(* IEC 61131-3 sources: deprecated-refusr-repo/GP/Main/samples (part 23) *)

(* ---- RND-EXPR_roust-surfs-pairs.st ---- *)
(*
This code implements a randomly grown symbolic expression:

xor(xor(!(xor(xor(IN32, (!(!((IN49 | (!(IN19))) & (!(IN28 & (xor(xor(IN18, IN20), IN24))))))) & ((xor(xor(IN13, IN1), !(xor(xor(xor(xor(!(IN32), IN20 & IN18), IN50 & IN1), (IN10 & IN17) & (IN11 & IN39)), true & IN1)))) | (xor(xor((!(IN35)) | IN42, !(IN44 | ((!(IN28)) | IN34))), (!((xor(xor(IN28, IN8), IN8)) & IN14)) | (!(xor(xor(xor(xor(IN16, IN9), IN43), xor(xor(IN30, IN9), IN40)), IN50 | IN28))))))), xor(xor((xor(xor(!(((!(IN18)) & (!(IN40))) & (IN28 & (!(IN19)))), IN7), (!((xor(xor(IN34, IN23), IN2)) & (xor(xor(IN27, IN44), IN31)))) | (!(xor(xor(!(IN25), IN8 & IN22), IN9))))) & (xor(xor(IN3, (!(IN42)) & (xor(xor(xor(xor(IN29 & IN50, IN38 | IN40), !(IN36)), IN40), (!(IN24)) & false))), (((!(IN11)) | (!(IN14))) | ((!(IN10)) | (IN36 & IN47))) | IN15)), (!(!(IN45))) & (xor(xor(IN31 | true, IN38), xor(xor(IN43, xor(xor(IN1, (IN12 & IN45) | (IN48 | IN6)), xor(xor(xor(xor(IN28, IN15), IN16), IN6), !(IN49)))), IN13 | ((xor(xor(IN45, IN5), IN32)) & (xor(xor(IN49, IN26), IN28))))))), !((!(IN43)) | (IN45 | (IN20 & (!(xor(xor(IN16, IN7), IN9))))))))), xor(xor((IN15 & ((!(xor(xor(!(xor(xor(IN18 | IN27, xor(xor(IN38, IN31), IN37)), !(IN3))), IN8 & (!(IN28 | IN17))), (xor(xor(IN17 | IN48, xor(xor(IN42, true), true)), IN31 | IN45)) | (IN25 | (!(IN12)))))) | ((!((xor(xor(!(IN16), IN16), xor(xor(IN32, IN22), IN35))) | IN22)) & ((!(xor(xor(IN8, xor(xor(IN18, IN44), IN32)), IN10 | IN3))) & (IN48 & (IN40 | (IN42 & IN27))))))) & IN10, ((!(!(xor(xor(IN3, IN47), (!(IN36 & IN49)) | ((xor(xor(IN42, IN21), IN34)) | (xor(xor(IN24, IN27), IN13))))))) | ((!(IN3)) & IN11)) & (!(((xor(xor(IN31 & IN15, ((!(IN49)) & (xor(xor(IN42, IN39), IN29))) & IN5), (IN7 | (IN32 | IN49)) & ((!(IN32)) | IN44))) & (!(!(!(IN47 & IN34))))) | (((true | (xor(xor(!(IN5), IN9 | IN38), !(IN46)))) | (!((IN37 | IN29) | (IN12 & IN37)))) | IN9)))), !((xor(xor(xor(xor(!(IN20), IN29 | IN30), (xor(xor(IN2, (IN21 & IN3) | (IN13 | IN7)), IN28)) | (xor(xor(IN44, IN21), (!(IN49)) & (!(IN44))))), xor(xor(xor(xor(xor(xor((!(IN48)) & (xor(xor(IN4, IN4), IN39)), (IN31 & IN45) & (IN44 | IN11)), IN5), IN42 & IN13), xor(xor(IN42, (xor(xor(IN14, IN11), IN43)) & IN1), true & (!(IN29)))), !(IN20)), true | (((xor(xor(IN15, IN17), IN17)) | IN20) | (!(!(IN29)))))), (!(IN1 | (xor(xor(IN14 & IN10, !(IN14)), IN21 & IN34)))) & IN17)) | ((IN1 & (xor(xor((!(IN2 & IN15)) | IN22, (!(IN21)) | (IN15 & IN29)), !(xor(xor(IN40, IN7 & IN9), IN31))))) & (((((IN44 & IN35) & (!(IN27))) | IN14) & (IN31 | ((!(IN25)) | (!(IN45))))) | (IN34 | (!((IN22 | IN16) & IN33)))))))), !(IN31 & ((!(xor(xor(((xor(xor(IN2 & IN9, IN28 & IN31), !(IN12))) | ((IN37 | IN35) | IN39)) | ((xor(xor(IN39 & IN49, IN2), IN26 | IN19)) | IN2), xor(xor((IN41 & (!(IN16))) & (xor(xor(!(IN33), IN12 & IN24), IN29 & IN35)), ((IN50 | IN17) & (IN41 & IN40)) | IN5), xor(xor(true, xor(xor(!(IN50), xor(xor(IN37, IN38), IN12)), !(IN47))), !(IN11 | IN42)))), IN42 | IN28))) | ((IN38 & IN43) & IN36))))

*)

FUNCTION_BLOCK F_CollectInput
  VAR_IN_OUT
      Data : ARRAY[1..50] OF BOOL;
  END_VAR
  VAR_INPUT
      TICK  : BOOL := 0;
      IN1   : BOOL := 0;
      IN2   : BOOL := 0;
      IN3   : BOOL := 0;
      IN4   : BOOL := 0;
      IN5   : BOOL := 0;
      RESET : BOOL := FALSE;
  END_VAR
  VAR_OUTPUT
      Finished : BOOL;
  END_VAR
  VAR
      j    : USINT := 1;
      tock : BOOL  := 0;
  END_VAR
  IF NOT RESET AND tock = NOT TICK THEN
      Data[j]   := IN1;
      Data[j+1] := IN2;
      Data[j+2] := IN3;
      Data[j+3] := IN4;
      Data[j+4] := IN5;
      j := j + 5;
      tock := TICK;
  ELSE
      j := 1;
      tock := 0;
  END_IF;
  Finished := (j > 50);
END_FUNCTION_BLOCK

PROGRAM Boiler
  VAR
    Data  : ARRAY[1..50] OF BOOL;
    Ready : BOOL;
    CollectInput : F_CollectInput;
  END_VAR
  VAR
    TICK     AT %IX1.0 : BOOL;
    IN1      AT %IX0.3 : BOOL;
    IN2      AT %IX0.4 : BOOL;
    IN3      AT %IX0.5 : BOOL;
    IN4      AT %IX0.6 : BOOL;
    IN5      AT %IX0.7 : BOOL;
    OutReady AT %QX0.0 : BOOL := FALSE;
    FeedNext AT %QX0.1 : BOOL := FALSE;
    Out      AT %QX0.2 : BOOL;
  END_VAR
  CollectInput(TICK:=TICK, IN1:=IN1, IN2:=IN2, IN3:=IN3, IN4:=IN4, IN5:=IN5);
  Ready := CollectInput.Finished;
  FeedNext := 1;
  IF Ready THEN
    Out := (((NOT ((Data[32] XOR ((NOT (NOT ((Data[49] OR (NOT Data[19])) AND (NOT (Data[28] AND ((Data[18] XOR Data[20]) XOR Data[24])))))) AND (((Data[13] XOR Data[1]) XOR (NOT (((((NOT Data[32]) XOR (Data[20] AND Data[18])) XOR (Data[50] AND Data[1])) XOR ((Data[10] AND Data[17]) AND (Data[11] AND Data[39]))) XOR (TRUE AND Data[1])))) OR ((((NOT Data[35]) OR Data[42]) XOR (NOT (Data[44] OR ((NOT Data[28]) OR Data[34])))) XOR ((NOT (((Data[28] XOR Data[8]) XOR Data[8]) AND Data[14])) OR (NOT ((((Data[16] XOR Data[9]) XOR Data[43]) XOR ((Data[30] XOR Data[9]) XOR Data[40])) XOR (Data[50] OR Data[28])))))))) XOR ((((((NOT (((NOT Data[18]) AND (NOT Data[40])) AND (Data[28] AND (NOT Data[19])))) XOR Data[7]) XOR ((NOT (((Data[34] XOR Data[23]) XOR Data[2]) AND ((Data[27] XOR Data[44]) XOR Data[31]))) OR (NOT (((NOT Data[25]) XOR (Data[8] AND Data[22])) XOR Data[9])))) AND ((Data[3] XOR ((NOT Data[42]) AND (((((Data[29] AND Data[50]) XOR (Data[38] OR Data[40])) XOR (NOT Data[36])) XOR Data[40]) XOR ((NOT Data[24]) AND FALSE)))) XOR ((((NOT Data[11]) OR (NOT Data[14])) OR ((NOT Data[10]) OR (Data[36] AND Data[47]))) OR Data[15]))) XOR ((NOT (NOT Data[45])) AND (((Data[31] OR TRUE) XOR Data[38]) XOR ((Data[43] XOR ((Data[1] XOR ((Data[12] AND Data[45]) OR (Data[48] OR Data[6]))) XOR ((((Data[28] XOR Data[15]) XOR Data[16]) XOR Data[6]) XOR (NOT Data[49])))) XOR (Data[13] OR (((Data[45] XOR Data[5]) XOR Data[32]) AND ((Data[49] XOR Data[26]) XOR Data[28]))))))) XOR (NOT ((NOT Data[43]) OR (Data[45] OR (Data[20] AND (NOT ((Data[16] XOR Data[7]) XOR Data[9]))))))))) XOR ((((Data[15] AND ((NOT (((NOT (((Data[18] OR Data[27]) XOR ((Data[38] XOR Data[31]) XOR Data[37])) XOR (NOT Data[3]))) XOR (Data[8] AND (NOT (Data[28] OR Data[17])))) XOR ((((Data[17] OR Data[48]) XOR ((Data[42] XOR TRUE) XOR TRUE)) XOR (Data[31] OR Data[45])) OR (Data[25] OR (NOT Data[12]))))) OR ((NOT ((((NOT Data[16]) XOR Data[16]) XOR ((Data[32] XOR Data[22]) XOR Data[35])) OR Data[22])) AND ((NOT ((Data[8] XOR ((Data[18] XOR Data[44]) XOR Data[32])) XOR (Data[10] OR Data[3]))) AND (Data[48] AND (Data[40] OR (Data[42] AND Data[27]))))))) AND Data[10]) XOR (((NOT (NOT ((Data[3] XOR Data[47]) XOR ((NOT (Data[36] AND Data[49])) OR (((Data[42] XOR Data[21]) XOR Data[34]) OR ((Data[24] XOR Data[27]) XOR Data[13])))))) OR ((NOT Data[3]) AND Data[11])) AND (NOT (((((Data[31] AND Data[15]) XOR (((NOT Data[49]) AND ((Data[42] XOR Data[39]) XOR Data[29])) AND Data[5])) XOR ((Data[7] OR (Data[32] OR Data[49])) AND ((NOT Data[32]) OR Data[44]))) AND (NOT (NOT (NOT (Data[47] AND Data[34]))))) OR (((TRUE OR (((NOT Data[5]) XOR (Data[9] OR Data[38])) XOR (NOT Data[46]))) OR (NOT ((Data[37] OR Data[29]) OR (Data[12] AND Data[37])))) OR Data[9]))))) XOR (NOT ((((((NOT Data[20]) XOR (Data[29] OR Data[30])) XOR (((Data[2] XOR ((Data[21] AND Data[3]) OR (Data[13] OR Data[7]))) XOR Data[28]) OR ((Data[44] XOR Data[21]) XOR ((NOT Data[49]) AND (NOT Data[44]))))) XOR ((((((((NOT Data[48]) AND ((Data[4] XOR Data[4]) XOR Data[39])) XOR ((Data[31] AND Data[45]) AND (Data[44] OR Data[11]))) XOR Data[5]) XOR (Data[42] AND Data[13])) XOR ((Data[42] XOR (((Data[14] XOR Data[11]) XOR Data[43]) AND Data[1])) XOR (TRUE AND (NOT Data[29])))) XOR (NOT Data[20])) XOR (TRUE OR ((((Data[15] XOR Data[17]) XOR Data[17]) OR Data[20]) OR (NOT (NOT Data[29])))))) XOR ((NOT (Data[1] OR (((Data[14] AND Data[10]) XOR (NOT Data[14])) XOR (Data[21] AND Data[34])))) AND Data[17])) OR ((Data[1] AND ((((NOT (Data[2] AND Data[15])) OR Data[22]) XOR ((NOT Data[21]) OR (Data[15] AND Data[29]))) XOR (NOT ((Data[40] XOR (Data[7] AND Data[9])) XOR Data[31])))) AND (((((Data[44] AND Data[35]) AND (NOT Data[27])) OR Data[14]) AND (Data[31] OR ((NOT Data[25]) OR (NOT Data[45])))) OR (Data[34] OR (NOT ((Data[22] OR Data[16]) AND Data[33]))))))))) XOR (NOT (Data[31] AND ((NOT (((((((Data[2] AND Data[9]) XOR (Data[28] AND Data[31])) XOR (NOT Data[12])) OR ((Data[37] OR Data[35]) OR Data[39])) OR ((((Data[39] AND Data[49]) XOR Data[2]) XOR (Data[26] OR Data[19])) OR Data[2])) XOR ((((Data[41] AND (NOT Data[16])) AND (((NOT Data[33]) XOR (Data[12] AND Data[24])) XOR (Data[29] AND Data[35]))) XOR (((Data[50] OR Data[17]) AND (Data[41] AND Data[40])) OR Data[5])) XOR ((TRUE XOR (((NOT Data[50]) XOR ((Data[37] XOR Data[38]) XOR Data[12])) XOR (NOT Data[47]))) XOR (NOT (Data[11] OR Data[42]))))) XOR (Data[42] OR Data[28]))) OR ((Data[38] AND Data[43]) AND Data[36])))));
    OutReady := 1;
    CollectInput(RESET:=TRUE);
  END_IF;
END_PROGRAM

CONFIGURATION Config0
  RESOURCE Res0 ON PLC
    TASK task0(INTERVAL := T#20ms,PRIORITY := 0);
    PROGRAM instance0 WITH task0 : Boiler;
  END_RESOURCE
END_CONFIGURATION

(* ---- RND-EXPR_sepal-sighs-minis.st ---- *)
(*
This code implements a randomly grown symbolic expression:

((xor(xor(!(IN17), IN3), IN42 & (!(!((!(xor(xor(IN42 & IN8, IN18), IN49))) | (!(IN32))))))) & ((!(!((IN47 | (IN12 & (xor(xor(!(IN9), IN41 & IN17), IN45)))) & (xor(xor(IN6 & (IN23 | (IN31 | IN44)), xor(xor((!(IN32)) & (!(IN23)), IN42 & (IN50 | IN34)), xor(xor(!(IN34), !(IN32)), IN15))), xor(xor(IN33, xor(xor(IN45 & IN5, IN11 & IN16), IN3 | IN4)), !(!(IN15)))))))) & (((xor(xor(((xor(xor(IN50 | IN14, IN46 & IN40), xor(xor(IN3, IN41), IN9))) & (IN22 & IN28)) | (xor(xor(IN41 | (IN26 & IN10), xor(xor(IN42 & IN12, xor(xor(IN32, IN46), IN35)), IN1 & IN11)), xor(xor(xor(xor(IN43, IN19), IN38), IN27 | IN21), !(IN10)))), !(xor(xor((xor(xor(IN7, IN50), IN1)) | IN6, (IN35 & IN3) | (!(IN28))), xor(xor(IN7 & IN16, IN37 | IN33), IN11)))), (!((!(IN25)) | (!(IN41)))) & ((!(IN33 & true)) & (!(!(IN5)))))) & (xor(xor(IN12, !(IN17)), (((!(IN28)) & (xor(xor(IN4, IN22), IN12))) | ((IN4 & IN38) & IN37)) | true))) | IN6))) & (xor(xor(!(IN24), xor(xor(!((xor(xor(IN48 | (!((IN17 & IN14) | IN31)), (xor(xor(true, xor(xor(xor(xor(IN16, IN16), IN17), !(IN23)), IN2)), (!(IN45)) | (xor(xor(IN31, IN48), IN25)))) & (!(xor(xor(IN6, IN41 & IN37), IN38)))), (IN26 | ((IN7 & IN2) | (IN17 | false))) & (xor(xor(IN42 & (IN28 | IN44), (IN16 & IN26) | (IN21 | IN13)), (IN11 & IN4) | (IN48 | IN47))))) & ((!(false & ((xor(xor(IN20, IN8), IN2)) | (IN36 & IN18)))) & IN47)), xor(xor(((false & (xor(xor(xor(xor(IN27 | IN30, xor(xor(IN23, IN27), IN7)), IN21), !(IN50)), (!(IN35)) & (xor(xor(IN21, IN7), IN17))))) | ((((IN9 | IN5) | (xor(xor(IN46, IN31), IN33))) | IN14) | IN32)) | (((!(IN19)) & IN21) & (!((!(IN44 & IN26)) | IN42))), xor(xor(!(IN34), (IN31 | (xor(xor(IN20, IN9), IN30))) | (xor(xor(IN21, xor(xor((IN29 | IN5) | (IN10 & IN14), xor(xor(IN41 & IN34, xor(xor(IN20, IN4), IN29)), IN29 & IN17)), IN39 | (IN7 & IN43))), ((!(IN40)) | IN50) | (!(IN17))))), xor(xor(xor(xor(IN31, IN24), ((IN30 | IN5) & (!(IN48))) | ((xor(xor(IN16, IN13), IN34)) & (!(IN16)))), (xor(xor(IN29 | IN25, xor(xor(xor(xor(IN20, IN40), IN9), IN26 | IN20), IN43 | IN32)), (xor(xor(IN35, IN6), IN33)) | (IN30 | IN7))) & (((true | IN15) | (IN46 | IN5)) | ((xor(xor(IN20, IN39), IN5)) | (IN48 | IN20)))), ((!(IN11 & IN1)) | ((xor(xor(IN5, IN25), IN49)) | (IN3 & IN43))) | (!(xor(xor(IN22, xor(xor(IN40, IN26), IN7)), xor(xor(IN10, IN10), IN44))))))), !(xor(xor(!(xor(xor((!(IN32)) | (xor(xor(IN28, IN4), IN11)), (IN7 | IN49) & (IN19 | IN17)), xor(xor(xor(xor(IN50, IN4), IN7), !(IN25)), !(IN10)))), (xor(xor(IN18 & (IN23 | IN36), xor(xor(IN36 | false, IN31 | IN19), IN15 & IN5)), !(IN41))) | (!(!(xor(xor(IN34, IN8), true))))), IN10 & (((IN39 & IN8) | (xor(xor(IN37, IN1), IN46))) | ((xor(xor(IN21, IN1), IN16)) | (false | IN1))))))), IN25 & (IN31 & (IN20 & IN46)))), IN38 | (!(IN32))))

*)

FUNCTION_BLOCK F_CollectInput
  VAR_IN_OUT
      Data : ARRAY[1..50] OF BOOL;
  END_VAR
  VAR_INPUT
      TICK  : BOOL := 0;
      IN1   : BOOL := 0;
      IN2   : BOOL := 0;
      IN3   : BOOL := 0;
      IN4   : BOOL := 0;
      IN5   : BOOL := 0;
      RESET : BOOL := FALSE;
  END_VAR
  VAR_OUTPUT
      Finished : BOOL;
  END_VAR
  VAR
      j    : USINT := 1;
      tock : BOOL  := 0;
  END_VAR
  IF NOT RESET AND tock = NOT TICK THEN
      Data[j]   := IN1;
      Data[j+1] := IN2;
      Data[j+2] := IN3;
      Data[j+3] := IN4;
      Data[j+4] := IN5;
      j := j + 5;
      tock := TICK;
  ELSE
      j := 1;
      tock := 0;
  END_IF;
  Finished := (j > 50);
END_FUNCTION_BLOCK

PROGRAM Boiler
  VAR
    Data  : ARRAY[1..50] OF BOOL;
    Ready : BOOL;
    CollectInput : F_CollectInput;
  END_VAR
  VAR
    TICK     AT %IX1.0 : BOOL;
    IN1      AT %IX0.3 : BOOL;
    IN2      AT %IX0.4 : BOOL;
    IN3      AT %IX0.5 : BOOL;
    IN4      AT %IX0.6 : BOOL;
    IN5      AT %IX0.7 : BOOL;
    OutReady AT %QX0.0 : BOOL := FALSE;
    FeedNext AT %QX0.1 : BOOL := FALSE;
    Out      AT %QX0.2 : BOOL;
  END_VAR
  CollectInput(TICK:=TICK, IN1:=IN1, IN2:=IN2, IN3:=IN3, IN4:=IN4, IN5:=IN5);
  Ready := CollectInput.Finished;
  FeedNext := 1;
  IF Ready THEN
    Out := (((((NOT Data[17]) XOR Data[3]) XOR (Data[42] AND (NOT (NOT ((NOT (((Data[42] AND Data[8]) XOR Data[18]) XOR Data[49])) OR (NOT Data[32])))))) AND ((NOT (NOT ((Data[47] OR (Data[12] AND (((NOT Data[9]) XOR (Data[41] AND Data[17])) XOR Data[45]))) AND (((Data[6] AND (Data[23] OR (Data[31] OR Data[44]))) XOR ((((NOT Data[32]) AND (NOT Data[23])) XOR (Data[42] AND (Data[50] OR Data[34]))) XOR (((NOT Data[34]) XOR (NOT Data[32])) XOR Data[15]))) XOR ((Data[33] XOR (((Data[45] AND Data[5]) XOR (Data[11] AND Data[16])) XOR (Data[3] OR Data[4]))) XOR (NOT (NOT Data[15]))))))) AND (((((((((Data[50] OR Data[14]) XOR (Data[46] AND Data[40])) XOR ((Data[3] XOR Data[41]) XOR Data[9])) AND (Data[22] AND Data[28])) OR (((Data[41] OR (Data[26] AND Data[10])) XOR (((Data[42] AND Data[12]) XOR ((Data[32] XOR Data[46]) XOR Data[35])) XOR (Data[1] AND Data[11]))) XOR ((((Data[43] XOR Data[19]) XOR Data[38]) XOR (Data[27] OR Data[21])) XOR (NOT Data[10])))) XOR (NOT (((((Data[7] XOR Data[50]) XOR Data[1]) OR Data[6]) XOR ((Data[35] AND Data[3]) OR (NOT Data[28]))) XOR (((Data[7] AND Data[16]) XOR (Data[37] OR Data[33])) XOR Data[11])))) XOR ((NOT ((NOT Data[25]) OR (NOT Data[41]))) AND ((NOT (Data[33] AND TRUE)) AND (NOT (NOT Data[5]))))) AND ((Data[12] XOR (NOT Data[17])) XOR ((((NOT Data[28]) AND ((Data[4] XOR Data[22]) XOR Data[12])) OR ((Data[4] AND Data[38]) AND Data[37])) OR TRUE))) OR Data[6]))) AND (((NOT Data[24]) XOR (((NOT ((((Data[48] OR (NOT ((Data[17] AND Data[14]) OR Data[31]))) XOR (((TRUE XOR ((((Data[16] XOR Data[16]) XOR Data[17]) XOR (NOT Data[23])) XOR Data[2])) XOR ((NOT Data[45]) OR ((Data[31] XOR Data[48]) XOR Data[25]))) AND (NOT ((Data[6] XOR (Data[41] AND Data[37])) XOR Data[38])))) XOR ((Data[26] OR ((Data[7] AND Data[2]) OR (Data[17] OR FALSE))) AND (((Data[42] AND (Data[28] OR Data[44])) XOR ((Data[16] AND Data[26]) OR (Data[21] OR Data[13]))) XOR ((Data[11] AND Data[4]) OR (Data[48] OR Data[47]))))) AND ((NOT (FALSE AND (((Data[20] XOR Data[8]) XOR Data[2]) OR (Data[36] AND Data[18])))) AND Data[47]))) XOR (((((FALSE AND (((((Data[27] OR Data[30]) XOR ((Data[23] XOR Data[27]) XOR Data[7])) XOR Data[21]) XOR (NOT Data[50])) XOR ((NOT Data[35]) AND ((Data[21] XOR Data[7]) XOR Data[17])))) OR ((((Data[9] OR Data[5]) OR ((Data[46] XOR Data[31]) XOR Data[33])) OR Data[14]) OR Data[32])) OR (((NOT Data[19]) AND Data[21]) AND (NOT ((NOT (Data[44] AND Data[26])) OR Data[42])))) XOR (((NOT Data[34]) XOR ((Data[31] OR ((Data[20] XOR Data[9]) XOR Data[30])) OR ((Data[21] XOR ((((Data[29] OR Data[5]) OR (Data[10] AND Data[14])) XOR (((Data[41] AND Data[34]) XOR ((Data[20] XOR Data[4]) XOR Data[29])) XOR (Data[29] AND Data[17]))) XOR (Data[39] OR (Data[7] AND Data[43])))) XOR (((NOT Data[40]) OR Data[50]) OR (NOT Data[17]))))) XOR ((((Data[31] XOR Data[24]) XOR (((Data[30] OR Data[5]) AND (NOT Data[48])) OR (((Data[16] XOR Data[13]) XOR Data[34]) AND (NOT Data[16])))) XOR ((((Data[29] OR Data[25]) XOR ((((Data[20] XOR Data[40]) XOR Data[9]) XOR (Data[26] OR Data[20])) XOR (Data[43] OR Data[32]))) XOR (((Data[35] XOR Data[6]) XOR Data[33]) OR (Data[30] OR Data[7]))) AND (((TRUE OR Data[15]) OR (Data[46] OR Data[5])) OR (((Data[20] XOR Data[39]) XOR Data[5]) OR (Data[48] OR Data[20]))))) XOR (((NOT (Data[11] AND Data[1])) OR (((Data[5] XOR Data[25]) XOR Data[49]) OR (Data[3] AND Data[43]))) OR (NOT ((Data[22] XOR ((Data[40] XOR Data[26]) XOR Data[7])) XOR ((Data[10] XOR Data[10]) XOR Data[44]))))))) XOR (NOT (((NOT ((((NOT Data[32]) OR ((Data[28] XOR Data[4]) XOR Data[11])) XOR ((Data[7] OR Data[49]) AND (Data[19] OR Data[17]))) XOR ((((Data[50] XOR Data[4]) XOR Data[7]) XOR (NOT Data[25])) XOR (NOT Data[10])))) XOR ((((Data[18] AND (Data[23] OR Data[36])) XOR (((Data[36] OR FALSE) XOR (Data[31] OR Data[19])) XOR (Data[15] AND Data[5]))) XOR (NOT Data[41])) OR (NOT (NOT ((Data[34] XOR Data[8]) XOR TRUE))))) XOR (Data[10] AND (((Data[39] AND Data[8]) OR ((Data[37] XOR Data[1]) XOR Data[46])) OR (((Data[21] XOR Data[1]) XOR Data[16]) OR (FALSE OR Data[1])))))))) XOR (Data[25] AND (Data[31] AND (Data[20] AND Data[46]))))) XOR (Data[38] OR (NOT Data[32]))));
    OutReady := 1;
    CollectInput(RESET:=TRUE);
  END_IF;
END_PROGRAM

CONFIGURATION Config0
  RESOURCE Res0 ON PLC
    TASK task0(INTERVAL := T#20ms,PRIORITY := 0);
    PROGRAM instance0 WITH task0 : Boiler;
  END_RESOURCE
END_CONFIGURATION

(* ---- RND-EXPR_sewed-hokey-cooch.st ---- *)
(*
This code implements a randomly grown symbolic expression:

!(((!(IN1)) | (xor(xor(!(IN4 | (!(xor(xor((!(IN21)) | (IN10 | IN34), (IN32 & IN39) & (xor(xor(IN33, IN21), IN30))), !(IN10 & IN16))))), !(!(!(xor(xor(IN12 & (!(IN27)), xor(xor(IN33 | IN30, IN41 & IN39), !(IN28))), IN32))))), xor(xor(!(!(IN49)), xor(xor((((IN3 & IN10) | (IN5 & IN27)) | IN6) & (IN43 | (xor(xor(IN8 | IN6, IN18 | IN20), IN22))), ((xor(xor(!(IN49), xor(xor(IN25, IN15), IN10)), xor(xor(IN36, IN47), IN50))) & false) | (!(xor(xor(!(IN13), IN25), xor(xor(IN8, IN43), IN45))))), IN44)), !(xor(xor(xor(xor((IN50 | IN36) | IN39, IN13), IN21), IN46 & IN31), IN9)))))) & (xor(xor(!((!(IN49)) | (xor(xor(!(IN31), IN49), (xor(xor(IN13, (xor(xor(IN6, IN49), IN32)) & (xor(xor(IN30, IN18), IN32))), IN42 | (IN13 | IN3))) & IN32))), ((!(xor(xor(xor(xor(IN31, IN16 | (!(IN20))), (true | IN11) | (IN30 & IN6)), ((xor(xor(IN5, IN18), IN47)) | (xor(xor(IN35, IN32), IN7))) & (!(IN35 | IN25))), (xor(xor(IN45 | IN27, !(IN16)), IN28 & IN24)) & ((IN12 | IN15) | (!(IN26)))))) & (!(IN14 & (((IN50 | IN36) & (!(IN18))) | (xor(xor(false, IN20 | IN26), IN25 | IN46)))))) & (!(IN16))), !((xor(xor((xor(xor((xor(xor(IN18, IN5), IN4)) & (IN10 | IN28), (IN14 | IN50) & (xor(xor(IN31, IN38), IN9))), (IN6 | IN10) | (IN46 | IN30))) | IN8, xor(xor((IN26 & (xor(xor(IN38, IN2), IN26))) & IN24, xor(xor(IN39, (xor(xor(IN4, IN26), IN46)) & (IN21 | IN23)), (IN46 | IN28) & (IN43 & IN9))), IN47)), (!((xor(xor(IN32, IN28), IN18)) & (IN11 & IN35))) & (((xor(xor(IN50, false), IN45)) & IN3) | (xor(xor(IN8, IN14 & IN13), IN48))))) | (((!(IN19)) | (IN26 & (!(!(IN22))))) & IN12)))))

*)

FUNCTION_BLOCK F_CollectInput
  VAR_IN_OUT
      Data : ARRAY[1..50] OF BOOL;
  END_VAR
  VAR_INPUT
      TICK  : BOOL := 0;
      IN1   : BOOL := 0;
      IN2   : BOOL := 0;
      IN3   : BOOL := 0;
      IN4   : BOOL := 0;
      IN5   : BOOL := 0;
      RESET : BOOL := FALSE;
  END_VAR
  VAR_OUTPUT
      Finished : BOOL;
  END_VAR
  VAR
      j    : USINT := 1;
      tock : BOOL  := 0;
  END_VAR
  IF NOT RESET AND tock = NOT TICK THEN
      Data[j]   := IN1;
      Data[j+1] := IN2;
      Data[j+2] := IN3;
      Data[j+3] := IN4;
      Data[j+4] := IN5;
      j := j + 5;
      tock := TICK;
  ELSE
      j := 1;
      tock := 0;
  END_IF;
  Finished := (j > 50);
END_FUNCTION_BLOCK

PROGRAM Boiler
  VAR
    Data  : ARRAY[1..50] OF BOOL;
    Ready : BOOL;
    CollectInput : F_CollectInput;
  END_VAR
  VAR
    TICK     AT %IX1.0 : BOOL;
    IN1      AT %IX0.3 : BOOL;
    IN2      AT %IX0.4 : BOOL;
    IN3      AT %IX0.5 : BOOL;
    IN4      AT %IX0.6 : BOOL;
    IN5      AT %IX0.7 : BOOL;
    OutReady AT %QX0.0 : BOOL := FALSE;
    FeedNext AT %QX0.1 : BOOL := FALSE;
    Out      AT %QX0.2 : BOOL;
  END_VAR
  CollectInput(TICK:=TICK, IN1:=IN1, IN2:=IN2, IN3:=IN3, IN4:=IN4, IN5:=IN5);
  Ready := CollectInput.Finished;
  FeedNext := 1;
  IF Ready THEN
    Out := (NOT (((NOT Data[1]) OR (((NOT (Data[4] OR (NOT ((((NOT Data[21]) OR (Data[10] OR Data[34])) XOR ((Data[32] AND Data[39]) AND ((Data[33] XOR Data[21]) XOR Data[30]))) XOR (NOT (Data[10] AND Data[16])))))) XOR (NOT (NOT (NOT (((Data[12] AND (NOT Data[27])) XOR (((Data[33] OR Data[30]) XOR (Data[41] AND Data[39])) XOR (NOT Data[28]))) XOR Data[32]))))) XOR (((NOT (NOT Data[49])) XOR ((((((Data[3] AND Data[10]) OR (Data[5] AND Data[27])) OR Data[6]) AND (Data[43] OR (((Data[8] OR Data[6]) XOR (Data[18] OR Data[20])) XOR Data[22]))) XOR (((((NOT Data[49]) XOR ((Data[25] XOR Data[15]) XOR Data[10])) XOR ((Data[36] XOR Data[47]) XOR Data[50])) AND FALSE) OR (NOT (((NOT Data[13]) XOR Data[25]) XOR ((Data[8] XOR Data[43]) XOR Data[45]))))) XOR Data[44])) XOR (NOT ((((((Data[50] OR Data[36]) OR Data[39]) XOR Data[13]) XOR Data[21]) XOR (Data[46] AND Data[31])) XOR Data[9]))))) AND (((NOT ((NOT Data[49]) OR (((NOT Data[31]) XOR Data[49]) XOR (((Data[13] XOR (((Data[6] XOR Data[49]) XOR Data[32]) AND ((Data[30] XOR Data[18]) XOR Data[32]))) XOR (Data[42] OR (Data[13] OR Data[3]))) AND Data[32])))) XOR (((NOT ((((Data[31] XOR (Data[16] OR (NOT Data[20]))) XOR ((TRUE OR Data[11]) OR (Data[30] AND Data[6]))) XOR ((((Data[5] XOR Data[18]) XOR Data[47]) OR ((Data[35] XOR Data[32]) XOR Data[7])) AND (NOT (Data[35] OR Data[25])))) XOR ((((Data[45] OR Data[27]) XOR (NOT Data[16])) XOR (Data[28] AND Data[24])) AND ((Data[12] OR Data[15]) OR (NOT Data[26]))))) AND (NOT (Data[14] AND (((Data[50] OR Data[36]) AND (NOT Data[18])) OR ((FALSE XOR (Data[20] OR Data[26])) XOR (Data[25] OR Data[46])))))) AND (NOT Data[16]))) XOR (NOT (((((((((Data[18] XOR Data[5]) XOR Data[4]) AND (Data[10] OR Data[28])) XOR ((Data[14] OR Data[50]) AND ((Data[31] XOR Data[38]) XOR Data[9]))) XOR ((Data[6] OR Data[10]) OR (Data[46] OR Data[30]))) OR Data[8]) XOR ((((Data[26] AND ((Data[38] XOR Data[2]) XOR Data[26])) AND Data[24]) XOR ((Data[39] XOR (((Data[4] XOR Data[26]) XOR Data[46]) AND (Data[21] OR Data[23]))) XOR ((Data[46] OR Data[28]) AND (Data[43] AND Data[9])))) XOR Data[47])) XOR ((NOT (((Data[32] XOR Data[28]) XOR Data[18]) AND (Data[11] AND Data[35]))) AND ((((Data[50] XOR FALSE) XOR Data[45]) AND Data[3]) OR ((Data[8] XOR (Data[14] AND Data[13])) XOR Data[48])))) OR (((NOT Data[19]) OR (Data[26] AND (NOT (NOT Data[22])))) AND Data[12]))))));
    OutReady := 1;
    CollectInput(RESET:=TRUE);
  END_IF;
END_PROGRAM

CONFIGURATION Config0
  RESOURCE Res0 ON PLC
    TASK task0(INTERVAL := T#20ms,PRIORITY := 0);
    PROGRAM instance0 WITH task0 : Boiler;
  END_RESOURCE
END_CONFIGURATION

(* ---- RND-EXPR_sisal-keens-dweeb.st ---- *)
(*
This code implements a randomly grown symbolic expression:

((IN8 & (xor(xor(xor(xor(((!(xor(xor(IN20 & IN27, IN16 & IN35), !(IN38)))) | (xor(xor(IN48, (xor(xor(IN13, IN11), IN50)) | (xor(xor(IN27, IN2), IN19))), xor(xor(IN10, xor(xor(IN3, IN44), IN33)), !(IN13))))) & ((((!(IN49)) | IN45) | ((xor(xor(IN37, IN11), IN42)) & (!(IN15)))) | ((IN38 & (false | IN44)) | ((xor(xor(IN48, IN7), IN31)) & (!(IN5))))), IN48), !((!(IN46)) | ((!(!(IN4))) | (!(IN23 | IN49))))), (!(xor(xor((IN49 & (!(IN6))) & IN43, xor(xor(IN45, !(IN11 & IN3)), (xor(xor(IN10, IN26), IN11)) & (IN38 & IN47))), IN10))) & ((xor(xor(xor(xor(xor(xor(IN44 | IN8, IN37), xor(xor(true, IN3), IN6)), !(IN43 & IN23)), IN6), (!(IN23 & IN33)) & (!(IN39 | IN20))), xor(xor((!(IN21)) & (IN28 | IN37), !(IN33 | IN4)), IN40))) | (!(((!(IN41)) & IN50) & ((xor(xor(IN17, IN41), IN2)) & (IN10 & IN29)))))), xor(xor(IN13, (xor(xor(!(xor(xor(!(IN25), IN30 & IN3), !(IN26))), xor(xor((IN34 | IN33) | (!(IN36)), !(IN43 | IN2)), xor(xor(IN10 & IN46, !(IN22)), xor(xor(IN44, IN37), IN16)))), xor(xor((xor(xor(IN36, IN11), IN27)) | (IN13 | IN50), (IN42 & IN34) & (IN5 & IN43)), xor(xor(IN35, !(IN35)), xor(xor(IN1, IN26), IN25))))) | (xor(xor(!(IN39), xor(xor(!(IN45 | IN21), (IN44 & IN4) & (IN15 & IN10)), !(xor(xor(IN22, IN31), IN43)))), xor(xor((xor(xor(IN15, IN44), IN15)) & (IN25 | IN26), xor(xor(IN20 & IN21, IN14 & IN13), !(IN20))), (IN50 | IN32) | (IN7 & IN7))))), (xor(xor(!((IN16 & IN46) & (xor(xor(IN50, IN17), IN23))), IN22 & ((!(IN22)) | true)), (!(xor(xor(IN30, IN23), IN12))) | (xor(xor(IN27 | IN25, xor(xor(IN32, IN20), IN47)), xor(xor(IN49, IN34), false))))) | (xor(xor(IN28, ((xor(xor(IN22, IN8), IN38)) | IN20) | (!(IN17 & IN39))), ((xor(xor(IN8, IN50), IN25)) & (IN25 & IN41)) | IN40)))))) | IN43) | (!(!(xor(xor(xor(xor(!(!(!((!(IN47)) | (xor(xor(IN48, IN32), IN40))))), xor(xor(xor(xor(IN26 & (IN36 & (IN50 | IN12)), ((IN19 & IN10) & IN42) | (xor(xor(xor(xor(IN48, IN40), IN26), IN37 & false), IN26 | IN44))), (IN23 | (IN47 | IN39)) & (xor(xor(IN31 | IN24, IN26 & IN6), !(IN11)))), !(IN22)), !(IN4))), IN18 | IN18), xor(xor(IN50, (xor(xor(xor(xor(xor(xor(IN38, IN39 | IN10), xor(xor(IN36, IN16), IN5)), !(IN43)), (xor(xor(IN43, IN20), IN44)) & (!(IN24))), ((xor(xor(IN27, IN1), IN9)) | (xor(xor(IN4, IN24), IN13))) & IN12), ((IN29 | IN47) | (!(IN32))) | IN1)) | (xor(xor(((IN41 | IN14) & (IN15 & IN9)) & IN9, (!(IN23)) | (xor(xor(IN13 | IN38, IN13), xor(xor(IN36, IN48), IN31)))), xor(xor((IN7 | IN11) | (!(IN34)), (!(IN34)) | (IN43 & IN1)), (IN49 | IN16) | (!(IN49)))))), xor(xor((((false | IN17) | (xor(xor(IN3, IN13), IN3))) | (!(IN16 & true))) | (IN1 | IN25), ((!(IN50)) & (!(IN36 & IN1))) | (!(!(xor(xor(IN48, IN46), IN35))))), xor(xor(IN19 & ((IN28 & IN49) & (IN43 | IN40)), IN14), (!(IN38 | IN6)) & IN50)))), IN48 & (xor(xor(((!(IN41)) | ((xor(xor(IN14, IN38), IN48)) & IN50)) & ((xor(xor(IN11, IN18 & IN7), IN7 | IN20)) | (IN8 & (xor(xor(IN8, IN23), IN20)))), xor(xor((xor(xor(IN26 & IN21, IN4 | IN14), xor(xor(IN31, false), IN18))) & (xor(xor(IN37, IN14 & IN47), xor(xor(IN14, IN8), IN37))), !((xor(xor(IN3, IN24), IN28)) & IN29)), (IN27 | (!(IN44))) & IN22)), (!(IN29)) | (!((!(IN36)) | (IN23 | IN34)))))))))

*)

FUNCTION_BLOCK F_CollectInput
  VAR_IN_OUT
      Data : ARRAY[1..50] OF BOOL;
  END_VAR
  VAR_INPUT
      TICK  : BOOL := 0;
      IN1   : BOOL := 0;
      IN2   : BOOL := 0;
      IN3   : BOOL := 0;
      IN4   : BOOL := 0;
      IN5   : BOOL := 0;
      RESET : BOOL := FALSE;
  END_VAR
  VAR_OUTPUT
      Finished : BOOL;
  END_VAR
  VAR
      j    : USINT := 1;
      tock : BOOL  := 0;
  END_VAR
  IF NOT RESET AND tock = NOT TICK THEN
      Data[j]   := IN1;
      Data[j+1] := IN2;
      Data[j+2] := IN3;
      Data[j+3] := IN4;
      Data[j+4] := IN5;
      j := j + 5;
      tock := TICK;
  ELSE
      j := 1;
      tock := 0;
  END_IF;
  Finished := (j > 50);
END_FUNCTION_BLOCK

PROGRAM Boiler
  VAR
    Data  : ARRAY[1..50] OF BOOL;
    Ready : BOOL;
    CollectInput : F_CollectInput;
  END_VAR
  VAR
    TICK     AT %IX1.0 : BOOL;
    IN1      AT %IX0.3 : BOOL;
    IN2      AT %IX0.4 : BOOL;
    IN3      AT %IX0.5 : BOOL;
    IN4      AT %IX0.6 : BOOL;
    IN5      AT %IX0.7 : BOOL;
    OutReady AT %QX0.0 : BOOL := FALSE;
    FeedNext AT %QX0.1 : BOOL := FALSE;
    Out      AT %QX0.2 : BOOL;
  END_VAR
  CollectInput(TICK:=TICK, IN1:=IN1, IN2:=IN2, IN3:=IN3, IN4:=IN4, IN5:=IN5);
  Ready := CollectInput.Finished;
  FeedNext := 1;
  IF Ready THEN
    Out := (((Data[8] AND (((((((NOT (((Data[20] AND Data[27]) XOR (Data[16] AND Data[35])) XOR (NOT Data[38]))) OR ((Data[48] XOR (((Data[13] XOR Data[11]) XOR Data[50]) OR ((Data[27] XOR Data[2]) XOR Data[19]))) XOR ((Data[10] XOR ((Data[3] XOR Data[44]) XOR Data[33])) XOR (NOT Data[13])))) AND ((((NOT Data[49]) OR Data[45]) OR (((Data[37] XOR Data[11]) XOR Data[42]) AND (NOT Data[15]))) OR ((Data[38] AND (FALSE OR Data[44])) OR (((Data[48] XOR Data[7]) XOR Data[31]) AND (NOT Data[5]))))) XOR Data[48]) XOR (NOT ((NOT Data[46]) OR ((NOT (NOT Data[4])) OR (NOT (Data[23] OR Data[49])))))) XOR ((NOT ((((Data[49] AND (NOT Data[6])) AND Data[43]) XOR ((Data[45] XOR (NOT (Data[11] AND Data[3]))) XOR (((Data[10] XOR Data[26]) XOR Data[11]) AND (Data[38] AND Data[47])))) XOR Data[10])) AND ((((((((Data[44] OR Data[8]) XOR Data[37]) XOR ((TRUE XOR Data[3]) XOR Data[6])) XOR (NOT (Data[43] AND Data[23]))) XOR Data[6]) XOR ((NOT (Data[23] AND Data[33])) AND (NOT (Data[39] OR Data[20])))) XOR ((((NOT Data[21]) AND (Data[28] OR Data[37])) XOR (NOT (Data[33] OR Data[4]))) XOR Data[40])) OR (NOT (((NOT Data[41]) AND Data[50]) AND (((Data[17] XOR Data[41]) XOR Data[2]) AND (Data[10] AND Data[29]))))))) XOR ((Data[13] XOR ((((NOT (((NOT Data[25]) XOR (Data[30] AND Data[3])) XOR (NOT Data[26]))) XOR ((((Data[34] OR Data[33]) OR (NOT Data[36])) XOR (NOT (Data[43] OR Data[2]))) XOR (((Data[10] AND Data[46]) XOR (NOT Data[22])) XOR ((Data[44] XOR Data[37]) XOR Data[16])))) XOR (((((Data[36] XOR Data[11]) XOR Data[27]) OR (Data[13] OR Data[50])) XOR ((Data[42] AND Data[34]) AND (Data[5] AND Data[43]))) XOR ((Data[35] XOR (NOT Data[35])) XOR ((Data[1] XOR Data[26]) XOR Data[25])))) OR (((NOT Data[39]) XOR (((NOT (Data[45] OR Data[21])) XOR ((Data[44] AND Data[4]) AND (Data[15] AND Data[10]))) XOR (NOT ((Data[22] XOR Data[31]) XOR Data[43])))) XOR (((((Data[15] XOR Data[44]) XOR Data[15]) AND (Data[25] OR Data[26])) XOR (((Data[20] AND Data[21]) XOR (Data[14] AND Data[13])) XOR (NOT Data[20]))) XOR ((Data[50] OR Data[32]) OR (Data[7] AND Data[7])))))) XOR ((((NOT ((Data[16] AND Data[46]) AND ((Data[50] XOR Data[17]) XOR Data[23]))) XOR (Data[22] AND ((NOT Data[22]) OR TRUE))) XOR ((NOT ((Data[30] XOR Data[23]) XOR Data[12])) OR (((Data[27] OR Data[25]) XOR ((Data[32] XOR Data[20]) XOR Data[47])) XOR ((Data[49] XOR Data[34]) XOR FALSE)))) OR ((Data[28] XOR ((((Data[22] XOR Data[8]) XOR Data[38]) OR Data[20]) OR (NOT (Data[17] AND Data[39])))) XOR ((((Data[8] XOR Data[50]) XOR Data[25]) AND (Data[25] AND Data[41])) OR Data[40])))))) OR Data[43]) OR (NOT (NOT (((((NOT (NOT (NOT ((NOT Data[47]) OR ((Data[48] XOR Data[32]) XOR Data[40]))))) XOR (((((Data[26] AND (Data[36] AND (Data[50] OR Data[12]))) XOR (((Data[19] AND Data[10]) AND Data[42]) OR ((((Data[48] XOR Data[40]) XOR Data[26]) XOR (Data[37] AND FALSE)) XOR (Data[26] OR Data[44])))) XOR ((Data[23] OR (Data[47] OR Data[39])) AND (((Data[31] OR Data[24]) XOR (Data[26] AND Data[6])) XOR (NOT Data[11])))) XOR (NOT Data[22])) XOR (NOT Data[4]))) XOR (Data[18] OR Data[18])) XOR ((Data[50] XOR (((((((Data[38] XOR (Data[39] OR Data[10])) XOR ((Data[36] XOR Data[16]) XOR Data[5])) XOR (NOT Data[43])) XOR (((Data[43] XOR Data[20]) XOR Data[44]) AND (NOT Data[24]))) XOR ((((Data[27] XOR Data[1]) XOR Data[9]) OR ((Data[4] XOR Data[24]) XOR Data[13])) AND Data[12])) XOR (((Data[29] OR Data[47]) OR (NOT Data[32])) OR Data[1])) OR (((((Data[41] OR Data[14]) AND (Data[15] AND Data[9])) AND Data[9]) XOR ((NOT Data[23]) OR (((Data[13] OR Data[38]) XOR Data[13]) XOR ((Data[36] XOR Data[48]) XOR Data[31])))) XOR ((((Data[7] OR Data[11]) OR (NOT Data[34])) XOR ((NOT Data[34]) OR (Data[43] AND Data[1]))) XOR ((Data[49] OR Data[16]) OR (NOT Data[49])))))) XOR ((((((FALSE OR Data[17]) OR ((Data[3] XOR Data[13]) XOR Data[3])) OR (NOT (Data[16] AND TRUE))) OR (Data[1] OR Data[25])) XOR (((NOT Data[50]) AND (NOT (Data[36] AND Data[1]))) OR (NOT (NOT ((Data[48] XOR Data[46]) XOR Data[35]))))) XOR (((Data[19] AND ((Data[28] AND Data[49]) AND (Data[43] OR Data[40]))) XOR Data[14]) XOR ((NOT (Data[38] OR Data[6])) AND Data[50]))))) XOR (Data[48] AND (((((NOT Data[41]) OR (((Data[14] XOR Data[38]) XOR Data[48]) AND Data[50])) AND (((Data[11] XOR (Data[18] AND Data[7])) XOR (Data[7] OR Data[20])) OR (Data[8] AND ((Data[8] XOR Data[23]) XOR Data[20])))) XOR ((((((Data[26] AND Data[21]) XOR (Data[4] OR Data[14])) XOR ((Data[31] XOR FALSE) XOR Data[18])) AND ((Data[37] XOR (Data[14] AND Data[47])) XOR ((Data[14] XOR Data[8]) XOR Data[37]))) XOR (NOT (((Data[3] XOR Data[24]) XOR Data[28]) AND Data[29]))) XOR ((Data[27] OR (NOT Data[44])) AND Data[22]))) XOR ((NOT Data[29]) OR (NOT ((NOT Data[36]) OR (Data[23] OR Data[34]))))))))));
    OutReady := 1;
    CollectInput(RESET:=TRUE);
  END_IF;
END_PROGRAM

CONFIGURATION Config0
  RESOURCE Res0 ON PLC
    TASK task0(INTERVAL := T#20ms,PRIORITY := 0);
    PROGRAM instance0 WITH task0 : Boiler;
  END_RESOURCE
END_CONFIGURATION

(* ---- RND-EXPR_slack-mayst-pearl.st ---- *)
(*
This code implements a randomly grown symbolic expression:

IN17 | (!(!((xor(xor(xor(xor(!(((IN42 | IN28) & IN28) | ((IN44 & IN38) | (xor(xor(IN20, IN19), IN29)))), xor(xor(!(xor(xor(IN18, IN32), IN1)), (xor(xor(!(IN28), IN23 | true), IN21 & IN35)) | (xor(xor(IN18 | IN17, IN20 & IN16), IN40 & IN14))), IN13)), xor(xor(xor(xor(IN41 & (!(IN16)), !(xor(xor(IN22, IN4), IN17))), IN6), ((IN31 & IN41) | (!(IN11))) & IN31), ((xor(xor(IN22, IN44), IN41)) & IN34) | ((xor(xor(IN15, IN11), IN36)) | IN35))), (!(xor(xor((IN11 & IN30) | (IN38 & false), !(xor(xor(IN41, IN7), IN16))), xor(xor(IN30 & IN43, !(IN24)), xor(xor(IN39, IN43), IN41))))) & ((xor(xor(xor(xor(!(IN23), !(IN26)), IN50), xor(xor(!(IN46), !(IN19)), IN3 & IN45)), IN18)) | (xor(xor(xor(xor(IN2 | IN38, IN7 & IN42), IN25), xor(xor(xor(xor(IN45, IN22), IN25), IN39 | IN11), xor(xor(IN39, false), IN22))), !(xor(xor(IN49, IN22), IN35)))))), xor(xor((!((!(IN26)) & (!(IN47)))) & (IN4 | ((IN20 & IN17) & IN25)), IN16), ((xor(xor(!(IN27), IN3), xor(xor(IN14, IN50), IN41))) | IN31) & (xor(xor(!(IN5 & IN37), (!(IN21)) | (xor(xor(IN22, IN34), IN26))), IN36))))) | (IN14 | ((IN6 & (xor(xor(IN41 | (IN46 & IN7), xor(xor(!(IN32), !(IN19)), xor(xor(IN6, IN15), IN15))), (xor(xor(IN7, IN12), IN31)) | IN24))) | (!(IN20)))))))

*)

FUNCTION_BLOCK F_CollectInput
  VAR_IN_OUT
      Data : ARRAY[1..50] OF BOOL;
  END_VAR
  VAR_INPUT
      TICK  : BOOL := 0;
      IN1   : BOOL := 0;
      IN2   : BOOL := 0;
      IN3   : BOOL := 0;
      IN4   : BOOL := 0;
      IN5   : BOOL := 0;
      RESET : BOOL := FALSE;
  END_VAR
  VAR_OUTPUT
      Finished : BOOL;
  END_VAR
  VAR
      j    : USINT := 1;
      tock : BOOL  := 0;
  END_VAR
  IF NOT RESET AND tock = NOT TICK THEN
      Data[j]   := IN1;
      Data[j+1] := IN2;
      Data[j+2] := IN3;
      Data[j+3] := IN4;
      Data[j+4] := IN5;
      j := j + 5;
      tock := TICK;
  ELSE
      j := 1;
      tock := 0;
  END_IF;
  Finished := (j > 50);
END_FUNCTION_BLOCK

PROGRAM Boiler
  VAR
    Data  : ARRAY[1..50] OF BOOL;
    Ready : BOOL;
    CollectInput : F_CollectInput;
  END_VAR
  VAR
    TICK     AT %IX1.0 : BOOL;
    IN1      AT %IX0.3 : BOOL;
    IN2      AT %IX0.4 : BOOL;
    IN3      AT %IX0.5 : BOOL;
    IN4      AT %IX0.6 : BOOL;
    IN5      AT %IX0.7 : BOOL;
    OutReady AT %QX0.0 : BOOL := FALSE;
    FeedNext AT %QX0.1 : BOOL := FALSE;
    Out      AT %QX0.2 : BOOL;
  END_VAR
  CollectInput(TICK:=TICK, IN1:=IN1, IN2:=IN2, IN3:=IN3, IN4:=IN4, IN5:=IN5);
  Ready := CollectInput.Finished;
  FeedNext := 1;
  IF Ready THEN
    Out := (Data[17] OR (NOT (NOT ((((((NOT (((Data[42] OR Data[28]) AND Data[28]) OR ((Data[44] AND Data[38]) OR ((Data[20] XOR Data[19]) XOR Data[29])))) XOR (((NOT ((Data[18] XOR Data[32]) XOR Data[1])) XOR ((((NOT Data[28]) XOR (Data[23] OR TRUE)) XOR (Data[21] AND Data[35])) OR (((Data[18] OR Data[17]) XOR (Data[20] AND Data[16])) XOR (Data[40] AND Data[14])))) XOR Data[13])) XOR (((((Data[41] AND (NOT Data[16])) XOR (NOT ((Data[22] XOR Data[4]) XOR Data[17]))) XOR Data[6]) XOR (((Data[31] AND Data[41]) OR (NOT Data[11])) AND Data[31])) XOR ((((Data[22] XOR Data[44]) XOR Data[41]) AND Data[34]) OR (((Data[15] XOR Data[11]) XOR Data[36]) OR Data[35])))) XOR ((NOT ((((Data[11] AND Data[30]) OR (Data[38] AND FALSE)) XOR (NOT ((Data[41] XOR Data[7]) XOR Data[16]))) XOR (((Data[30] AND Data[43]) XOR (NOT Data[24])) XOR ((Data[39] XOR Data[43]) XOR Data[41])))) AND ((((((NOT Data[23]) XOR (NOT Data[26])) XOR Data[50]) XOR (((NOT Data[46]) XOR (NOT Data[19])) XOR (Data[3] AND Data[45]))) XOR Data[18]) OR (((((Data[2] OR Data[38]) XOR (Data[7] AND Data[42])) XOR Data[25]) XOR ((((Data[45] XOR Data[22]) XOR Data[25]) XOR (Data[39] OR Data[11])) XOR ((Data[39] XOR FALSE) XOR Data[22]))) XOR (NOT ((Data[49] XOR Data[22]) XOR Data[35])))))) XOR ((((NOT ((NOT Data[26]) AND (NOT Data[47]))) AND (Data[4] OR ((Data[20] AND Data[17]) AND Data[25]))) XOR Data[16]) XOR (((((NOT Data[27]) XOR Data[3]) XOR ((Data[14] XOR Data[50]) XOR Data[41])) OR Data[31]) AND (((NOT (Data[5] AND Data[37])) XOR ((NOT Data[21]) OR ((Data[22] XOR Data[34]) XOR Data[26]))) XOR Data[36])))) OR (Data[14] OR ((Data[6] AND (((Data[41] OR (Data[46] AND Data[7])) XOR (((NOT Data[32]) XOR (NOT Data[19])) XOR ((Data[6] XOR Data[15]) XOR Data[15]))) XOR (((Data[7] XOR Data[12]) XOR Data[31]) OR Data[24]))) OR (NOT Data[20])))))));
    OutReady := 1;
    CollectInput(RESET:=TRUE);
  END_IF;
END_PROGRAM

CONFIGURATION Config0
  RESOURCE Res0 ON PLC
    TASK task0(INTERVAL := T#20ms,PRIORITY := 0);
    PROGRAM instance0 WITH task0 : Boiler;
  END_RESOURCE
END_CONFIGURATION

(* ---- RND-EXPR_slyer-tutus-acing.st ---- *)
(*
This code implements a randomly grown symbolic expression:

IN41 & IN9

*)

FUNCTION_BLOCK F_CollectInput
  VAR_IN_OUT
      Data : ARRAY[1..50] OF BOOL;
  END_VAR
  VAR_INPUT
      TICK  : BOOL := 0;
      IN1   : BOOL := 0;
      IN2   : BOOL := 0;
      IN3   : BOOL := 0;
      IN4   : BOOL := 0;
      IN5   : BOOL := 0;
      RESET : BOOL := FALSE;
  END_VAR
  VAR_OUTPUT
      Finished : BOOL;
  END_VAR
  VAR
      j    : USINT := 1;
      tock : BOOL  := 0;
  END_VAR
  IF NOT RESET AND tock = NOT TICK THEN
      Data[j]   := IN1;
      Data[j+1] := IN2;
      Data[j+2] := IN3;
      Data[j+3] := IN4;
      Data[j+4] := IN5;
      j := j + 5;
      tock := TICK;
  ELSE
      j := 1;
      tock := 0;
  END_IF;
  Finished := (j > 50);
END_FUNCTION_BLOCK

PROGRAM Boiler
  VAR
    Data  : ARRAY[1..50] OF BOOL;
    Ready : BOOL;
    CollectInput : F_CollectInput;
  END_VAR
  VAR
    TICK     AT %IX1.0 : BOOL;
    IN1      AT %IX0.3 : BOOL;
    IN2      AT %IX0.4 : BOOL;
    IN3      AT %IX0.5 : BOOL;
    IN4      AT %IX0.6 : BOOL;
    IN5      AT %IX0.7 : BOOL;
    OutReady AT %QX0.0 : BOOL := FALSE;
    FeedNext AT %QX0.1 : BOOL := FALSE;
    Out      AT %QX0.2 : BOOL;
  END_VAR
  CollectInput(TICK:=TICK, IN1:=IN1, IN2:=IN2, IN3:=IN3, IN4:=IN4, IN5:=IN5);
  Ready := CollectInput.Finished;
  FeedNext := 1;
  IF Ready THEN
    Out := (Data[41] AND Data[9]);
    OutReady := 1;
    CollectInput(RESET:=TRUE);
  END_IF;
END_PROGRAM

CONFIGURATION Config0
  RESOURCE Res0 ON PLC
    TASK task0(INTERVAL := T#20ms,PRIORITY := 0);
    PROGRAM instance0 WITH task0 : Boiler;
  END_RESOURCE
END_CONFIGURATION

(* ---- RND-EXPR_snowy-guava-upend.st ---- *)
(*
This code implements a randomly grown symbolic expression:

(((((xor(xor((((IN14 | IN26) & (xor(xor(IN30, IN38), IN29))) | (xor(xor(IN43 | IN33, !(IN21)), IN49 | IN20))) & ((xor(xor(!(IN35), IN36), IN43 | IN5)) & (xor(xor(IN25 | IN20, IN28), !(IN27)))), (!(IN29)) | (!(true | (xor(xor(IN14, IN30), IN3))))), IN13)) | IN18) & ((xor(xor(xor(xor(IN43, !(IN44)), IN27), (!((!(IN48)) | false)) | (((!(IN39)) & (!(IN38))) | ((xor(xor(IN39, IN38), IN15)) & (xor(xor(IN18, IN2), IN41))))), (xor(xor(xor(xor(IN49 & IN31, xor(xor(IN13, IN22), IN6)), IN4 | IN40), (IN3 | IN27) | (!(IN6))), (xor(xor(IN22, IN8), IN42)) & (!(IN42)))) | ((xor(xor(xor(xor(IN12, IN36), IN50), !(IN14)), IN17 & IN37)) & true))) | true)) & (!(xor(xor((xor(xor(xor(xor(xor(xor(IN24 | IN1, IN3), IN17), xor(xor(IN50 | IN18, IN19), xor(xor(IN29, IN28), IN4))), (IN18 | false) | IN25), ((!(IN15)) & (!(IN2))) & IN4), xor(xor(IN33, (IN44 & IN37) & (xor(xor(IN49, IN7), IN25))), IN18))) & ((true & (!(IN11 & IN43))) & (((IN32 & IN13) & (xor(xor(IN12, IN19), false))) & true)), xor(xor((xor(xor((false | IN32) | (!(IN14)), (!(IN12)) & (xor(xor(IN49, IN4), true))), IN34)) | IN15, xor(xor(IN15, ((xor(xor(IN41, IN12), IN20)) | (xor(xor(IN21, IN44), IN18))) & (xor(xor(IN33 & IN12, IN25), xor(xor(IN1, IN19), true)))), xor(xor((IN49 | IN9) & (IN31 & false), !(IN49 | IN19)), (xor(xor(IN13, IN7), IN4)) | (true & IN34)))), xor(xor(xor(xor(IN15, (IN36 & IN11) & (xor(xor(IN46, IN33), IN2))), (xor(xor(IN29, IN36), false)) & (IN24 & IN12)), !(xor(xor(false & IN10, IN15), xor(xor(IN25, IN11), IN19)))), !(!(!(IN22)))))), IN14)))) & ((xor(xor(IN33 & IN5, xor(xor((!(xor(xor(xor(xor(!(IN34), !(IN15)), !(IN35)), !(IN7 | IN43)), xor(xor(!(IN45), IN23 | IN36), IN33 & IN5)))) & IN42, !(IN14)), (!(!(!(xor(xor(IN24, IN40), IN46))))) | IN22)), xor(xor(((((IN14 | IN48) | (xor(xor(IN38, IN48), IN19))) | IN42) | (((xor(xor(IN10, IN38), IN50)) | IN28) & (!(!(IN40))))) & IN30, IN41), ((!((IN11 & IN11) | (xor(xor(IN38, IN32), IN19)))) & ((!(IN44 & IN44)) | ((xor(xor(IN37, IN46), IN40)) & (!(IN19))))) & ((!(xor(xor(IN46, xor(xor(IN39, IN2), IN24)), xor(xor(IN1, IN43), IN50)))) & (((xor(xor(IN25, IN2), IN29)) | (IN34 & IN12)) & ((!(IN2)) & (xor(xor(IN14, IN33), IN13)))))))) & ((((((IN10 | (true | IN33)) & ((xor(xor(IN18, IN28), IN25)) & (!(IN25)))) & ((xor(xor(!(IN36), true | IN1), IN20)) & ((xor(xor(IN26, IN12), IN37)) | (false & IN15)))) & (((xor(xor(xor(xor(IN31, IN27), IN42), IN40 & IN2), IN42 & IN24)) & (xor(xor(IN47 | IN36, !(IN29)), IN2 | IN41))) & IN42)) | (xor(xor(xor(xor(!(!(IN9 & IN36)), !(xor(xor(IN16, IN28), IN32 | true))), ((xor(xor(IN10, IN24), IN46)) | (!(IN45))) & (!(IN37 & IN12))), (xor(xor(xor(xor(xor(xor(IN6, IN13), IN48), IN32 & IN7), xor(xor(IN34, IN19), IN46)), IN47), IN14 & (xor(xor(IN23, IN44), IN42)))) | IN35), (((IN8 & false) & (IN14 & IN20)) & IN19) | IN39))) & IN18))) | ((IN44 & true) & ((xor(xor((!(!(IN2 | ((xor(xor(IN32, IN15), IN7)) | (xor(xor(IN30, IN15), IN20)))))) & IN48, (xor(xor(((!(IN37)) & (!(xor(xor(IN36, IN13), IN21)))) & (IN7 & IN39), (!(IN13)) & (xor(xor(!(!(IN7)), IN34), false | (IN6 & IN16)))), (((IN41 & IN45) & (IN28 | IN39)) | (!(IN15 & IN38))) & (xor(xor(IN36, (IN48 | IN18) & (IN18 & IN20)), (xor(xor(IN47, IN26), IN11)) | (!(IN27)))))) & IN12), IN20)) | (((xor(xor(IN40, xor(xor(((IN7 & IN24) | (xor(xor(IN32, IN26), IN16))) | IN23, xor(xor(IN39 & (IN45 | IN19), xor(xor(xor(xor(IN41, IN17), IN4), xor(xor(IN6, IN46), IN22)), false & IN3)), (xor(xor(IN22, IN17), IN47)) | (!(IN15)))), !((xor(xor(IN25, IN5), IN24)) | (IN3 | IN29)))), (IN3 & (!(IN43))) & IN21)) & ((!(xor(xor((xor(xor(IN32, IN39), IN15)) & (!(IN21)), (IN37 | IN20) & (!(IN31))), xor(xor(IN25, IN28 & IN16), IN4 | IN17)))) & (!((xor(xor(xor(xor(IN31, IN25), IN5), xor(xor(IN1, IN10), IN50)), !(IN18))) | ((!(IN18)) | IN34))))) | (IN33 | ((!(((IN23 & IN13) & (IN3 | IN11)) & ((xor(xor(IN6, IN14), IN29)) | (IN20 | IN44)))) | (!(IN24 | ((xor(xor(IN28, IN29), IN10)) & (!(IN27))))))))))

*)

FUNCTION_BLOCK F_CollectInput
  VAR_IN_OUT
      Data : ARRAY[1..50] OF BOOL;
  END_VAR
  VAR_INPUT
      TICK  : BOOL := 0;
      IN1   : BOOL := 0;
      IN2   : BOOL := 0;
      IN3   : BOOL := 0;
      IN4   : BOOL := 0;
      IN5   : BOOL := 0;
      RESET : BOOL := FALSE;
  END_VAR
  VAR_OUTPUT
      Finished : BOOL;
  END_VAR
  VAR
      j    : USINT := 1;
      tock : BOOL  := 0;
  END_VAR
  IF NOT RESET AND tock = NOT TICK THEN
      Data[j]   := IN1;
      Data[j+1] := IN2;
      Data[j+2] := IN3;
      Data[j+3] := IN4;
      Data[j+4] := IN5;
      j := j + 5;
      tock := TICK;
  ELSE
      j := 1;
      tock := 0;
  END_IF;
  Finished := (j > 50);
END_FUNCTION_BLOCK

PROGRAM Boiler
  VAR
    Data  : ARRAY[1..50] OF BOOL;
    Ready : BOOL;
    CollectInput : F_CollectInput;
  END_VAR
  VAR
    TICK     AT %IX1.0 : BOOL;
    IN1      AT %IX0.3 : BOOL;
    IN2      AT %IX0.4 : BOOL;
    IN3      AT %IX0.5 : BOOL;
    IN4      AT %IX0.6 : BOOL;
    IN5      AT %IX0.7 : BOOL;
    OutReady AT %QX0.0 : BOOL := FALSE;
    FeedNext AT %QX0.1 : BOOL := FALSE;
    Out      AT %QX0.2 : BOOL;
  END_VAR
  CollectInput(TICK:=TICK, IN1:=IN1, IN2:=IN2, IN3:=IN3, IN4:=IN4, IN5:=IN5);
  Ready := CollectInput.Finished;
  FeedNext := 1;
  IF Ready THEN
    Out := (((((((((((Data[14] OR Data[26]) AND ((Data[30] XOR Data[38]) XOR Data[29])) OR (((Data[43] OR Data[33]) XOR (NOT Data[21])) XOR (Data[49] OR Data[20]))) AND ((((NOT Data[35]) XOR Data[36]) XOR (Data[43] OR Data[5])) AND (((Data[25] OR Data[20]) XOR Data[28]) XOR (NOT Data[27])))) XOR ((NOT Data[29]) OR (NOT (TRUE OR ((Data[14] XOR Data[30]) XOR Data[3]))))) XOR Data[13]) OR Data[18]) AND (((((Data[43] XOR (NOT Data[44])) XOR Data[27]) XOR ((NOT ((NOT Data[48]) OR FALSE)) OR (((NOT Data[39]) AND (NOT Data[38])) OR (((Data[39] XOR Data[38]) XOR Data[15]) AND ((Data[18] XOR Data[2]) XOR Data[41]))))) XOR ((((((Data[49] AND Data[31]) XOR ((Data[13] XOR Data[22]) XOR Data[6])) XOR (Data[4] OR Data[40])) XOR ((Data[3] OR Data[27]) OR (NOT Data[6]))) XOR (((Data[22] XOR Data[8]) XOR Data[42]) AND (NOT Data[42]))) OR (((((Data[12] XOR Data[36]) XOR Data[50]) XOR (NOT Data[14])) XOR (Data[17] AND Data[37])) AND TRUE))) OR TRUE)) AND (NOT ((((((((((Data[24] OR Data[1]) XOR Data[3]) XOR Data[17]) XOR (((Data[50] OR Data[18]) XOR Data[19]) XOR ((Data[29] XOR Data[28]) XOR Data[4]))) XOR ((Data[18] OR FALSE) OR Data[25])) XOR (((NOT Data[15]) AND (NOT Data[2])) AND Data[4])) XOR ((Data[33] XOR ((Data[44] AND Data[37]) AND ((Data[49] XOR Data[7]) XOR Data[25]))) XOR Data[18])) AND ((TRUE AND (NOT (Data[11] AND Data[43]))) AND (((Data[32] AND Data[13]) AND ((Data[12] XOR Data[19]) XOR FALSE)) AND TRUE))) XOR (((((((FALSE OR Data[32]) OR (NOT Data[14])) XOR ((NOT Data[12]) AND ((Data[49] XOR Data[4]) XOR TRUE))) XOR Data[34]) OR Data[15]) XOR ((Data[15] XOR ((((Data[41] XOR Data[12]) XOR Data[20]) OR ((Data[21] XOR Data[44]) XOR Data[18])) AND (((Data[33] AND Data[12]) XOR Data[25]) XOR ((Data[1] XOR Data[19]) XOR TRUE)))) XOR ((((Data[49] OR Data[9]) AND (Data[31] AND FALSE)) XOR (NOT (Data[49] OR Data[19]))) XOR (((Data[13] XOR Data[7]) XOR Data[4]) OR (TRUE AND Data[34]))))) XOR ((((Data[15] XOR ((Data[36] AND Data[11]) AND ((Data[46] XOR Data[33]) XOR Data[2]))) XOR (((Data[29] XOR Data[36]) XOR FALSE) AND (Data[24] AND Data[12]))) XOR (NOT (((FALSE AND Data[10]) XOR Data[15]) XOR ((Data[25] XOR Data[11]) XOR Data[19])))) XOR (NOT (NOT (NOT Data[22])))))) XOR Data[14]))) AND ((((Data[33] AND Data[5]) XOR ((((NOT (((((NOT Data[34]) XOR (NOT Data[15])) XOR (NOT Data[35])) XOR (NOT (Data[7] OR Data[43]))) XOR (((NOT Data[45]) XOR (Data[23] OR Data[36])) XOR (Data[33] AND Data[5])))) AND Data[42]) XOR (NOT Data[14])) XOR ((NOT (NOT (NOT ((Data[24] XOR Data[40]) XOR Data[46])))) OR Data[22]))) XOR (((((((Data[14] OR Data[48]) OR ((Data[38] XOR Data[48]) XOR Data[19])) OR Data[42]) OR ((((Data[10] XOR Data[38]) XOR Data[50]) OR Data[28]) AND (NOT (NOT Data[40])))) AND Data[30]) XOR Data[41]) XOR (((NOT ((Data[11] AND Data[11]) OR ((Data[38] XOR Data[32]) XOR Data[19]))) AND ((NOT (Data[44] AND Data[44])) OR (((Data[37] XOR Data[46]) XOR Data[40]) AND (NOT Data[19])))) AND ((NOT ((Data[46] XOR ((Data[39] XOR Data[2]) XOR Data[24])) XOR ((Data[1] XOR Data[43]) XOR Data[50]))) AND ((((Data[25] XOR Data[2]) XOR Data[29]) OR (Data[34] AND Data[12])) AND ((NOT Data[2]) AND ((Data[14] XOR Data[33]) XOR Data[13]))))))) AND ((((((Data[10] OR (TRUE OR Data[33])) AND (((Data[18] XOR Data[28]) XOR Data[25]) AND (NOT Data[25]))) AND ((((NOT Data[36]) XOR (TRUE OR Data[1])) XOR Data[20]) AND (((Data[26] XOR Data[12]) XOR Data[37]) OR (FALSE AND Data[15])))) AND ((((((Data[31] XOR Data[27]) XOR Data[42]) XOR (Data[40] AND Data[2])) XOR (Data[42] AND Data[24])) AND (((Data[47] OR Data[36]) XOR (NOT Data[29])) XOR (Data[2] OR Data[41]))) AND Data[42])) OR (((((NOT (NOT (Data[9] AND Data[36]))) XOR (NOT ((Data[16] XOR Data[28]) XOR (Data[32] OR TRUE)))) XOR ((((Data[10] XOR Data[24]) XOR Data[46]) OR (NOT Data[45])) AND (NOT (Data[37] AND Data[12])))) XOR (((((((Data[6] XOR Data[13]) XOR Data[48]) XOR (Data[32] AND Data[7])) XOR ((Data[34] XOR Data[19]) XOR Data[46])) XOR Data[47]) XOR (Data[14] AND ((Data[23] XOR Data[44]) XOR Data[42]))) OR Data[35])) XOR ((((Data[8] AND FALSE) AND (Data[14] AND Data[20])) AND Data[19]) OR Data[39]))) AND Data[18]))) OR ((Data[44] AND TRUE) AND (((((NOT (NOT (Data[2] OR (((Data[32] XOR Data[15]) XOR Data[7]) OR ((Data[30] XOR Data[15]) XOR Data[20]))))) AND Data[48]) XOR ((((((NOT Data[37]) AND (NOT ((Data[36] XOR Data[13]) XOR Data[21]))) AND (Data[7] AND Data[39])) XOR ((NOT Data[13]) AND (((NOT (NOT Data[7])) XOR Data[34]) XOR (FALSE OR (Data[6] AND Data[16]))))) XOR ((((Data[41] AND Data[45]) AND (Data[28] OR Data[39])) OR (NOT (Data[15] AND Data[38]))) AND ((Data[36] XOR ((Data[48] OR Data[18]) AND (Data[18] AND Data[20]))) XOR (((Data[47] XOR Data[26]) XOR Data[11]) OR (NOT Data[27]))))) AND Data[12])) XOR Data[20]) OR ((((Data[40] XOR (((((Data[7] AND Data[24]) OR ((Data[32] XOR Data[26]) XOR Data[16])) OR Data[23]) XOR (((Data[39] AND (Data[45] OR Data[19])) XOR ((((Data[41] XOR Data[17]) XOR Data[4]) XOR ((Data[6] XOR Data[46]) XOR Data[22])) XOR (FALSE AND Data[3]))) XOR (((Data[22] XOR Data[17]) XOR Data[47]) OR (NOT Data[15])))) XOR (NOT (((Data[25] XOR Data[5]) XOR Data[24]) OR (Data[3] OR Data[29]))))) XOR ((Data[3] AND (NOT Data[43])) AND Data[21])) AND ((NOT (((((Data[32] XOR Data[39]) XOR Data[15]) AND (NOT Data[21])) XOR ((Data[37] OR Data[20]) AND (NOT Data[31]))) XOR ((Data[25] XOR (Data[28] AND Data[16])) XOR (Data[4] OR Data[17])))) AND (NOT (((((Data[31] XOR Data[25]) XOR Data[5]) XOR ((Data[1] XOR Data[10]) XOR Data[50])) XOR (NOT Data[18])) OR ((NOT Data[18]) OR Data[34]))))) OR (Data[33] OR ((NOT (((Data[23] AND Data[13]) AND (Data[3] OR Data[11])) AND (((Data[6] XOR Data[14]) XOR Data[29]) OR (Data[20] OR Data[44])))) OR (NOT (Data[24] OR (((Data[28] XOR Data[29]) XOR Data[10]) AND (NOT Data[27]))))))))));
    OutReady := 1;
    CollectInput(RESET:=TRUE);
  END_IF;
END_PROGRAM

CONFIGURATION Config0
  RESOURCE Res0 ON PLC
    TASK task0(INTERVAL := T#20ms,PRIORITY := 0);
    PROGRAM instance0 WITH task0 : Boiler;
  END_RESOURCE
END_CONFIGURATION

(* ---- RND-EXPR_souls-kirks-linty.st ---- *)
(*
This code implements a randomly grown symbolic expression:

!((IN49 & (!((!(xor(xor(!(IN22 | (IN41 | IN43)), (!(IN35 & IN45)) | (!(IN31 & IN19))), (xor(xor(IN19 | IN38, IN23), IN36 & IN43)) & ((IN20 | IN36) | (IN29 | IN25))))) & (((((IN8 | IN23) | IN36) & ((!(IN1)) & IN50)) & (!(xor(xor(IN22 & IN34, IN21), IN29 & IN35)))) & (xor(xor(IN49 | (xor(xor(!(IN23), !(IN35)), IN10 & IN32)), (xor(xor(IN36, IN45 & IN19), !(IN16))) | (!(!(IN39)))), (xor(xor(xor(xor(IN43, IN46), IN50), IN32), !(IN48))) & IN17)))))) | ((xor(xor(xor(xor(xor(xor(IN37 | (!(!(IN47))), IN2), (((xor(xor(IN13, IN9), IN5)) & (IN37 | IN2)) | ((IN47 & IN30) | (IN14 | IN47))) & (xor(xor(!(IN25 | IN6), IN5), (IN46 & IN32) & (IN14 | IN49)))), !(!((xor(xor(!(IN41), IN1), xor(xor(IN20, IN32), IN5))) | (!(false | IN15))))), xor(xor(!(((IN41 | IN5) & (IN31 | IN34)) & (xor(xor(xor(xor(IN42, IN28), IN26), xor(xor(IN31, IN48), IN22)), !(IN36)))), ((xor(xor(IN22 | IN3, false | IN19), IN22 | IN10)) & ((xor(xor(IN5, IN38), IN13)) | (IN33 & IN25))) & (IN9 | (IN3 | (xor(xor(IN47, IN3), IN32))))), xor(xor(((IN19 & IN42) & (IN25 & IN35)) | (IN21 & (!(IN48))), false | (xor(xor(!(IN30), !(IN46)), IN34))), !((IN19 & IN26) | (xor(xor(IN45, IN3), IN18)))))), xor(xor(IN25, IN50), !(!(xor(xor(xor(xor(!(IN46), IN7 | IN20), !(IN34)), (!(IN18)) | (IN7 & IN5)), (IN38 | IN27) | (IN35 & IN3)))))), xor(xor(!((IN44 & (!(IN14))) | (((xor(xor(IN31, IN33), IN31)) | (!(IN23))) & ((IN20 | IN5) & (!(IN39))))), IN18), xor(xor(IN38, xor(xor(!(!(!(IN48))), ((IN32 & IN8) | (IN35 | IN22)) & ((IN18 | IN40) & true)), IN41)), IN26)))) & IN31))

*)

FUNCTION_BLOCK F_CollectInput
  VAR_IN_OUT
      Data : ARRAY[1..50] OF BOOL;
  END_VAR
  VAR_INPUT
      TICK  : BOOL := 0;
      IN1   : BOOL := 0;
      IN2   : BOOL := 0;
      IN3   : BOOL := 0;
      IN4   : BOOL := 0;
      IN5   : BOOL := 0;
      RESET : BOOL := FALSE;
  END_VAR
  VAR_OUTPUT
      Finished : BOOL;
  END_VAR
  VAR
      j    : USINT := 1;
      tock : BOOL  := 0;
  END_VAR
  IF NOT RESET AND tock = NOT TICK THEN
      Data[j]   := IN1;
      Data[j+1] := IN2;
      Data[j+2] := IN3;
      Data[j+3] := IN4;
      Data[j+4] := IN5;
      j := j + 5;
      tock := TICK;
  ELSE
      j := 1;
      tock := 0;
  END_IF;
  Finished := (j > 50);
END_FUNCTION_BLOCK

PROGRAM Boiler
  VAR
    Data  : ARRAY[1..50] OF BOOL;
    Ready : BOOL;
    CollectInput : F_CollectInput;
  END_VAR
  VAR
    TICK     AT %IX1.0 : BOOL;
    IN1      AT %IX0.3 : BOOL;
    IN2      AT %IX0.4 : BOOL;
    IN3      AT %IX0.5 : BOOL;
    IN4      AT %IX0.6 : BOOL;
    IN5      AT %IX0.7 : BOOL;
    OutReady AT %QX0.0 : BOOL := FALSE;
    FeedNext AT %QX0.1 : BOOL := FALSE;
    Out      AT %QX0.2 : BOOL;
  END_VAR
  CollectInput(TICK:=TICK, IN1:=IN1, IN2:=IN2, IN3:=IN3, IN4:=IN4, IN5:=IN5);
  Ready := CollectInput.Finished;
  FeedNext := 1;
  IF Ready THEN
    Out := (NOT ((Data[49] AND (NOT ((NOT (((NOT (Data[22] OR (Data[41] OR Data[43]))) XOR ((NOT (Data[35] AND Data[45])) OR (NOT (Data[31] AND Data[19])))) XOR ((((Data[19] OR Data[38]) XOR Data[23]) XOR (Data[36] AND Data[43])) AND ((Data[20] OR Data[36]) OR (Data[29] OR Data[25]))))) AND (((((Data[8] OR Data[23]) OR Data[36]) AND ((NOT Data[1]) AND Data[50])) AND (NOT (((Data[22] AND Data[34]) XOR Data[21]) XOR (Data[29] AND Data[35])))) AND (((Data[49] OR (((NOT Data[23]) XOR (NOT Data[35])) XOR (Data[10] AND Data[32]))) XOR (((Data[36] XOR (Data[45] AND Data[19])) XOR (NOT Data[16])) OR (NOT (NOT Data[39])))) XOR (((((Data[43] XOR Data[46]) XOR Data[50]) XOR Data[32]) XOR (NOT Data[48])) AND Data[17])))))) OR ((((((((Data[37] OR (NOT (NOT Data[47]))) XOR Data[2]) XOR (((((Data[13] XOR Data[9]) XOR Data[5]) AND (Data[37] OR Data[2])) OR ((Data[47] AND Data[30]) OR (Data[14] OR Data[47]))) AND (((NOT (Data[25] OR Data[6])) XOR Data[5]) XOR ((Data[46] AND Data[32]) AND (Data[14] OR Data[49]))))) XOR (NOT (NOT ((((NOT Data[41]) XOR Data[1]) XOR ((Data[20] XOR Data[32]) XOR Data[5])) OR (NOT (FALSE OR Data[15])))))) XOR (((NOT (((Data[41] OR Data[5]) AND (Data[31] OR Data[34])) AND ((((Data[42] XOR Data[28]) XOR Data[26]) XOR ((Data[31] XOR Data[48]) XOR Data[22])) XOR (NOT Data[36])))) XOR (((((Data[22] OR Data[3]) XOR (FALSE OR Data[19])) XOR (Data[22] OR Data[10])) AND (((Data[5] XOR Data[38]) XOR Data[13]) OR (Data[33] AND Data[25]))) AND (Data[9] OR (Data[3] OR ((Data[47] XOR Data[3]) XOR Data[32]))))) XOR (((((Data[19] AND Data[42]) AND (Data[25] AND Data[35])) OR (Data[21] AND (NOT Data[48]))) XOR (FALSE OR (((NOT Data[30]) XOR (NOT Data[46])) XOR Data[34]))) XOR (NOT ((Data[19] AND Data[26]) OR ((Data[45] XOR Data[3]) XOR Data[18])))))) XOR ((Data[25] XOR Data[50]) XOR (NOT (NOT (((((NOT Data[46]) XOR (Data[7] OR Data[20])) XOR (NOT Data[34])) XOR ((NOT Data[18]) OR (Data[7] AND Data[5]))) XOR ((Data[38] OR Data[27]) OR (Data[35] AND Data[3]))))))) XOR (((NOT ((Data[44] AND (NOT Data[14])) OR ((((Data[31] XOR Data[33]) XOR Data[31]) OR (NOT Data[23])) AND ((Data[20] OR Data[5]) AND (NOT Data[39]))))) XOR Data[18]) XOR ((Data[38] XOR (((NOT (NOT (NOT Data[48]))) XOR (((Data[32] AND Data[8]) OR (Data[35] OR Data[22])) AND ((Data[18] OR Data[40]) AND TRUE))) XOR Data[41])) XOR Data[26]))) AND Data[31])));
    OutReady := 1;
    CollectInput(RESET:=TRUE);
  END_IF;
END_PROGRAM

CONFIGURATION Config0
  RESOURCE Res0 ON PLC
    TASK task0(INTERVAL := T#20ms,PRIORITY := 0);
    PROGRAM instance0 WITH task0 : Boiler;
  END_RESOURCE
END_CONFIGURATION

(* ---- RND-EXPR_spits-coven-beryl.st ---- *)
(*
This code implements a randomly grown symbolic expression:

!(!((((!(!((IN26 | (IN14 | IN47)) | ((IN43 & IN29) & (IN9 & IN8))))) | (((!(IN30 & IN26)) | ((xor(xor(IN9 & IN4, xor(xor(IN26, IN10), false)), xor(xor(IN41, IN12), IN33))) | ((xor(xor(IN25, IN41), IN50)) | (IN36 & IN45)))) | (!(xor(xor(IN43, !(IN26 & IN49)), xor(xor(!(IN41), IN20), !(IN35))))))) | (((xor(xor(xor(xor((IN25 & IN40) | (!(IN50)), xor(xor(IN1 | IN36, IN48 & IN11), !(IN9))), xor(xor(xor(xor(IN29, IN24), IN16), IN4), IN32 & IN26)), (!(IN25)) & (IN10 & IN22)), !((!(IN26)) | (!(IN19))))) & (xor(xor(IN41, xor(xor(xor(xor(IN45, IN33), IN10 & IN46), IN37), (!(IN28)) | (!(IN26)))), IN49))) & IN18)) & (xor(xor(((!(xor(xor((IN47 | IN27) | (IN10 | IN23), (!(IN36)) & false), true | (!(IN44))))) | (xor(xor(xor(xor(xor(xor(IN35 & IN39, xor(xor(IN21, IN41), IN43)), !(IN2)), (IN5 & IN41) | (IN29 | false)), (IN8 | IN23) & IN30), (xor(xor(!(IN18), xor(xor(IN36, IN27), IN17)), IN21 | true)) & IN1), (!(IN37 & true)) | ((IN5 & IN1) & IN14)))) & IN7, (!(!(IN35))) | (((xor(xor((IN45 & IN3) | (!(IN10)), (xor(xor(IN8, IN19), IN50)) | (IN35 & IN12)), true | IN46)) | (((IN43 | IN4) | (!(IN20))) & ((IN3 | IN22) & (!(IN41))))) & (xor(xor((xor(xor(xor(xor(IN40, IN44), IN16), IN20), !(IN19))) & IN31, (xor(xor(IN40 & IN6, xor(xor(IN49, IN42), IN24)), !(IN33))) & (xor(xor(!(IN31), xor(xor(IN6, IN28), IN4)), xor(xor(IN15, IN42), IN47)))), (IN18 & (IN12 & IN17)) | (!(IN6 | IN21)))))), (!(xor(xor(IN27, (!(!(IN39))) & (xor(xor(!(IN37), IN42 & IN9), xor(xor(IN17, IN41), IN39)))), xor(xor(IN48, (xor(xor(IN40, IN7), IN9)) & (IN17 & IN6)), IN49)))) & ((!(xor(xor(IN3 & (!(IN18)), !(IN19 | IN43)), !(xor(xor(IN34, IN48), IN28))))) & ((!(xor(xor(IN29 | IN13, !(IN23)), !(IN1)))) & (xor(xor((IN44 | IN32) & (xor(xor(IN34, IN3), IN24)), IN43), (IN25 | IN11) | (xor(xor(IN14, IN26), IN44))))))))))

*)

FUNCTION_BLOCK F_CollectInput
  VAR_IN_OUT
      Data : ARRAY[1..50] OF BOOL;
  END_VAR
  VAR_INPUT
      TICK  : BOOL := 0;
      IN1   : BOOL := 0;
      IN2   : BOOL := 0;
      IN3   : BOOL := 0;
      IN4   : BOOL := 0;
      IN5   : BOOL := 0;
      RESET : BOOL := FALSE;
  END_VAR
  VAR_OUTPUT
      Finished : BOOL;
  END_VAR
  VAR
      j    : USINT := 1;
      tock : BOOL  := 0;
  END_VAR
  IF NOT RESET AND tock = NOT TICK THEN
      Data[j]   := IN1;
      Data[j+1] := IN2;
      Data[j+2] := IN3;
      Data[j+3] := IN4;
      Data[j+4] := IN5;
      j := j + 5;
      tock := TICK;
  ELSE
      j := 1;
      tock := 0;
  END_IF;
  Finished := (j > 50);
END_FUNCTION_BLOCK

PROGRAM Boiler
  VAR
    Data  : ARRAY[1..50] OF BOOL;
    Ready : BOOL;
    CollectInput : F_CollectInput;
  END_VAR
  VAR
    TICK     AT %IX1.0 : BOOL;
    IN1      AT %IX0.3 : BOOL;
    IN2      AT %IX0.4 : BOOL;
    IN3      AT %IX0.5 : BOOL;
    IN4      AT %IX0.6 : BOOL;
    IN5      AT %IX0.7 : BOOL;
    OutReady AT %QX0.0 : BOOL := FALSE;
    FeedNext AT %QX0.1 : BOOL := FALSE;
    Out      AT %QX0.2 : BOOL;
  END_VAR
  CollectInput(TICK:=TICK, IN1:=IN1, IN2:=IN2, IN3:=IN3, IN4:=IN4, IN5:=IN5);
  Ready := CollectInput.Finished;
  FeedNext := 1;
  IF Ready THEN
    Out := (NOT (NOT ((((NOT (NOT ((Data[26] OR (Data[14] OR Data[47])) OR ((Data[43] AND Data[29]) AND (Data[9] AND Data[8]))))) OR (((NOT (Data[30] AND Data[26])) OR ((((Data[9] AND Data[4]) XOR ((Data[26] XOR Data[10]) XOR FALSE)) XOR ((Data[41] XOR Data[12]) XOR Data[33])) OR (((Data[25] XOR Data[41]) XOR Data[50]) OR (Data[36] AND Data[45])))) OR (NOT ((Data[43] XOR (NOT (Data[26] AND Data[49]))) XOR (((NOT Data[41]) XOR Data[20]) XOR (NOT Data[35])))))) OR ((((((((Data[25] AND Data[40]) OR (NOT Data[50])) XOR (((Data[1] OR Data[36]) XOR (Data[48] AND Data[11])) XOR (NOT Data[9]))) XOR ((((Data[29] XOR Data[24]) XOR Data[16]) XOR Data[4]) XOR (Data[32] AND Data[26]))) XOR ((NOT Data[25]) AND (Data[10] AND Data[22]))) XOR (NOT ((NOT Data[26]) OR (NOT Data[19])))) AND ((Data[41] XOR ((((Data[45] XOR Data[33]) XOR (Data[10] AND Data[46])) XOR Data[37]) XOR ((NOT Data[28]) OR (NOT Data[26])))) XOR Data[49])) AND Data[18])) AND (((((NOT ((((Data[47] OR Data[27]) OR (Data[10] OR Data[23])) XOR ((NOT Data[36]) AND FALSE)) XOR (TRUE OR (NOT Data[44])))) OR (((((((Data[35] AND Data[39]) XOR ((Data[21] XOR Data[41]) XOR Data[43])) XOR (NOT Data[2])) XOR ((Data[5] AND Data[41]) OR (Data[29] OR FALSE))) XOR ((Data[8] OR Data[23]) AND Data[30])) XOR ((((NOT Data[18]) XOR ((Data[36] XOR Data[27]) XOR Data[17])) XOR (Data[21] OR TRUE)) AND Data[1])) XOR ((NOT (Data[37] AND TRUE)) OR ((Data[5] AND Data[1]) AND Data[14])))) AND Data[7]) XOR ((NOT (NOT Data[35])) OR ((((((Data[45] AND Data[3]) OR (NOT Data[10])) XOR (((Data[8] XOR Data[19]) XOR Data[50]) OR (Data[35] AND Data[12]))) XOR (TRUE OR Data[46])) OR (((Data[43] OR Data[4]) OR (NOT Data[20])) AND ((Data[3] OR Data[22]) AND (NOT Data[41])))) AND (((((((Data[40] XOR Data[44]) XOR Data[16]) XOR Data[20]) XOR (NOT Data[19])) AND Data[31]) XOR ((((Data[40] AND Data[6]) XOR ((Data[49] XOR Data[42]) XOR Data[24])) XOR (NOT Data[33])) AND (((NOT Data[31]) XOR ((Data[6] XOR Data[28]) XOR Data[4])) XOR ((Data[15] XOR Data[42]) XOR Data[47])))) XOR ((Data[18] AND (Data[12] AND Data[17])) OR (NOT (Data[6] OR Data[21]))))))) XOR ((NOT ((Data[27] XOR ((NOT (NOT Data[39])) AND (((NOT Data[37]) XOR (Data[42] AND Data[9])) XOR ((Data[17] XOR Data[41]) XOR Data[39])))) XOR ((Data[48] XOR (((Data[40] XOR Data[7]) XOR Data[9]) AND (Data[17] AND Data[6]))) XOR Data[49]))) AND ((NOT (((Data[3] AND (NOT Data[18])) XOR (NOT (Data[19] OR Data[43]))) XOR (NOT ((Data[34] XOR Data[48]) XOR Data[28])))) AND ((NOT (((Data[29] OR Data[13]) XOR (NOT Data[23])) XOR (NOT Data[1]))) AND ((((Data[44] OR Data[32]) AND ((Data[34] XOR Data[3]) XOR Data[24])) XOR Data[43]) XOR ((Data[25] OR Data[11]) OR ((Data[14] XOR Data[26]) XOR Data[44]))))))))));
    OutReady := 1;
    CollectInput(RESET:=TRUE);
  END_IF;
END_PROGRAM

CONFIGURATION Config0
  RESOURCE Res0 ON PLC
    TASK task0(INTERVAL := T#20ms,PRIORITY := 0);
    PROGRAM instance0 WITH task0 : Boiler;
  END_RESOURCE
END_CONFIGURATION

(* ---- RND-EXPR_start-licks-barmy.st ---- *)
(*
This code implements a randomly grown symbolic expression:

((((xor(xor(xor(xor((xor(xor(!(!(IN8)), IN19 | (IN35 | IN37)), !(IN12))) | IN7, ((xor(xor(IN20 | IN2, xor(xor(IN27, IN40), IN7)), IN16)) & (!(IN17 | IN17))) & ((xor(xor(IN45, IN7), xor(xor(IN1, IN44), IN25))) & (!(xor(xor(IN14, IN43), IN36))))), true), (xor(xor(IN15, !(IN44)), xor(xor((!(IN11)) & (xor(xor(IN49, IN16), IN8)), (IN32 | IN48) & (IN42 | IN18)), xor(xor(!(IN22), xor(xor(IN48, IN32), IN36)), !(IN17))))) | ((!((!(IN34)) & (IN32 | IN4))) | (xor(xor((IN39 | IN26) & IN24, IN5), xor(xor(IN6, IN27 | IN11), IN7 | IN20))))), !(!(!((IN30 & IN50) & (xor(xor(IN19, IN1), IN19))))))) | (xor(xor((!(IN26 | IN34)) | (IN49 | (xor(xor(IN18 & (IN36 | IN36), (IN49 | IN44) & IN50), IN41))), xor(xor(xor(xor((IN4 & IN44) | (!(!(IN49))), xor(xor((xor(xor(IN22, IN46), IN16)) & (!(IN50)), IN35), (IN48 | IN37) | (IN31 & IN24))), IN28 & IN22), !(IN39 | (xor(xor(!(IN40), IN22 & IN9), IN45 | IN44)))), (IN37 & (xor(xor(IN11 | IN6, IN1 & IN33), IN48 | IN8))) | (((xor(xor(IN13, IN21), IN23)) & (IN8 & IN13)) & (!(xor(xor(IN19, IN11), IN41)))))), (IN16 & (((xor(xor(IN48, IN5), IN44)) | IN8) & ((xor(xor(IN8, IN45), IN50)) | (xor(xor(false, IN6), IN41))))) | ((xor(xor((xor(xor(IN4, IN16), IN7)) | (!(IN40)), xor(xor(IN41 | IN45, IN30 & IN33), xor(xor(IN22, IN47), IN1))), xor(xor(!(IN1), IN10 & IN6), xor(xor(IN42, IN48), IN2)))) & IN37)))) | (((!(((!(IN2 & IN39)) & ((!(IN27)) & (IN32 | IN14))) & ((!(IN7 & IN12)) | IN26))) & (IN18 & ((!((IN12 & IN32) & (xor(xor(false, IN10), IN24)))) & true))) & (xor(xor((!(IN9 | (!(IN47)))) | (IN43 & IN17), IN35), IN20)))) | (((IN42 & (xor(xor(((!(xor(xor(IN9, IN3), IN36))) & ((IN18 & IN39) | (true & IN42))) | (!((IN25 & IN25) | IN46)), xor(xor(!(!(IN4 & IN44)), IN45), (!(!(IN47))) | ((!(IN44)) | (xor(xor(IN35, IN38), IN27))))), !(xor(xor(IN27, IN27), !(IN33 | IN35)))))) & (IN32 | (xor(xor((xor(xor(IN36, (IN37 & IN8) & (!(IN37))), IN9)) | (IN22 & ((IN15 & IN45) | (!(IN12)))), (((IN38 & IN46) & (IN45 & IN49)) & (IN2 & (xor(xor(IN46, IN25), IN24)))) & ((IN8 | (IN10 & IN25)) | (xor(xor(!(IN46), IN19 & IN11), !(IN20))))), ((xor(xor(xor(xor(IN22, IN26), IN31), IN7 | IN40), IN21)) & (!(!(IN32)))) | (((IN40 | IN1) & IN32) | ((IN37 | IN35) & (IN1 & IN45))))))) | (xor(xor((IN25 | IN42) & ((xor(xor((xor(xor(IN35, !(IN28)), IN12 | IN17)) | IN25, ((xor(xor(IN3, IN2), IN25)) & (IN32 | IN9)) & (xor(xor(IN33 & IN43, !(IN37)), IN28 & IN2))), false)) & IN30), IN36), IN6)))) & (!(!(IN43)))

*)

FUNCTION_BLOCK F_CollectInput
  VAR_IN_OUT
      Data : ARRAY[1..50] OF BOOL;
  END_VAR
  VAR_INPUT
      TICK  : BOOL := 0;
      IN1   : BOOL := 0;
      IN2   : BOOL := 0;
      IN3   : BOOL := 0;
      IN4   : BOOL := 0;
      IN5   : BOOL := 0;
      RESET : BOOL := FALSE;
  END_VAR
  VAR_OUTPUT
      Finished : BOOL;
  END_VAR
  VAR
      j    : USINT := 1;
      tock : BOOL  := 0;
  END_VAR
  IF NOT RESET AND tock = NOT TICK THEN
      Data[j]   := IN1;
      Data[j+1] := IN2;
      Data[j+2] := IN3;
      Data[j+3] := IN4;
      Data[j+4] := IN5;
      j := j + 5;
      tock := TICK;
  ELSE
      j := 1;
      tock := 0;
  END_IF;
  Finished := (j > 50);
END_FUNCTION_BLOCK

PROGRAM Boiler
  VAR
    Data  : ARRAY[1..50] OF BOOL;
    Ready : BOOL;
    CollectInput : F_CollectInput;
  END_VAR
  VAR
    TICK     AT %IX1.0 : BOOL;
    IN1      AT %IX0.3 : BOOL;
    IN2      AT %IX0.4 : BOOL;
    IN3      AT %IX0.5 : BOOL;
    IN4      AT %IX0.6 : BOOL;
    IN5      AT %IX0.7 : BOOL;
    OutReady AT %QX0.0 : BOOL := FALSE;
    FeedNext AT %QX0.1 : BOOL := FALSE;
    Out      AT %QX0.2 : BOOL;
  END_VAR
  CollectInput(TICK:=TICK, IN1:=IN1, IN2:=IN2, IN3:=IN3, IN4:=IN4, IN5:=IN5);
  Ready := CollectInput.Finished;
  FeedNext := 1;
  IF Ready THEN
    Out := ((((((((((((NOT (NOT Data[8])) XOR (Data[19] OR (Data[35] OR Data[37]))) XOR (NOT Data[12])) OR Data[7]) XOR (((((Data[20] OR Data[2]) XOR ((Data[27] XOR Data[40]) XOR Data[7])) XOR Data[16]) AND (NOT (Data[17] OR Data[17]))) AND (((Data[45] XOR Data[7]) XOR ((Data[1] XOR Data[44]) XOR Data[25])) AND (NOT ((Data[14] XOR Data[43]) XOR Data[36]))))) XOR TRUE) XOR (((Data[15] XOR (NOT Data[44])) XOR ((((NOT Data[11]) AND ((Data[49] XOR Data[16]) XOR Data[8])) XOR ((Data[32] OR Data[48]) AND (Data[42] OR Data[18]))) XOR (((NOT Data[22]) XOR ((Data[48] XOR Data[32]) XOR Data[36])) XOR (NOT Data[17])))) OR ((NOT ((NOT Data[34]) AND (Data[32] OR Data[4]))) OR ((((Data[39] OR Data[26]) AND Data[24]) XOR Data[5]) XOR ((Data[6] XOR (Data[27] OR Data[11])) XOR (Data[7] OR Data[20])))))) XOR (NOT (NOT (NOT ((Data[30] AND Data[50]) AND ((Data[19] XOR Data[1]) XOR Data[19])))))) OR ((((NOT (Data[26] OR Data[34])) OR (Data[49] OR (((Data[18] AND (Data[36] OR Data[36])) XOR ((Data[49] OR Data[44]) AND Data[50])) XOR Data[41]))) XOR ((((((Data[4] AND Data[44]) OR (NOT (NOT Data[49]))) XOR (((((Data[22] XOR Data[46]) XOR Data[16]) AND (NOT Data[50])) XOR Data[35]) XOR ((Data[48] OR Data[37]) OR (Data[31] AND Data[24])))) XOR (Data[28] AND Data[22])) XOR (NOT (Data[39] OR (((NOT Data[40]) XOR (Data[22] AND Data[9])) XOR (Data[45] OR Data[44]))))) XOR ((Data[37] AND (((Data[11] OR Data[6]) XOR (Data[1] AND Data[33])) XOR (Data[48] OR Data[8]))) OR ((((Data[13] XOR Data[21]) XOR Data[23]) AND (Data[8] AND Data[13])) AND (NOT ((Data[19] XOR Data[11]) XOR Data[41])))))) XOR ((Data[16] AND ((((Data[48] XOR Data[5]) XOR Data[44]) OR Data[8]) AND (((Data[8] XOR Data[45]) XOR Data[50]) OR ((FALSE XOR Data[6]) XOR Data[41])))) OR ((((((Data[4] XOR Data[16]) XOR Data[7]) OR (NOT Data[40])) XOR (((Data[41] OR Data[45]) XOR (Data[30] AND Data[33])) XOR ((Data[22] XOR Data[47]) XOR Data[1]))) XOR (((NOT Data[1]) XOR (Data[10] AND Data[6])) XOR ((Data[42] XOR Data[48]) XOR Data[2]))) AND Data[37])))) OR (((NOT (((NOT (Data[2] AND Data[39])) AND ((NOT Data[27]) AND (Data[32] OR Data[14]))) AND ((NOT (Data[7] AND Data[12])) OR Data[26]))) AND (Data[18] AND ((NOT ((Data[12] AND Data[32]) AND ((FALSE XOR Data[10]) XOR Data[24]))) AND TRUE))) AND ((((NOT (Data[9] OR (NOT Data[47]))) OR (Data[43] AND Data[17])) XOR Data[35]) XOR Data[20]))) OR (((Data[42] AND (((((NOT ((Data[9] XOR Data[3]) XOR Data[36])) AND ((Data[18] AND Data[39]) OR (TRUE AND Data[42]))) OR (NOT ((Data[25] AND Data[25]) OR Data[46]))) XOR (((NOT (NOT (Data[4] AND Data[44]))) XOR Data[45]) XOR ((NOT (NOT Data[47])) OR ((NOT Data[44]) OR ((Data[35] XOR Data[38]) XOR Data[27]))))) XOR (NOT ((Data[27] XOR Data[27]) XOR (NOT (Data[33] OR Data[35])))))) AND (Data[32] OR (((((Data[36] XOR ((Data[37] AND Data[8]) AND (NOT Data[37]))) XOR Data[9]) OR (Data[22] AND ((Data[15] AND Data[45]) OR (NOT Data[12])))) XOR ((((Data[38] AND Data[46]) AND (Data[45] AND Data[49])) AND (Data[2] AND ((Data[46] XOR Data[25]) XOR Data[24]))) AND ((Data[8] OR (Data[10] AND Data[25])) OR (((NOT Data[46]) XOR (Data[19] AND Data[11])) XOR (NOT Data[20]))))) XOR ((((((Data[22] XOR Data[26]) XOR Data[31]) XOR (Data[7] OR Data[40])) XOR Data[21]) AND (NOT (NOT Data[32]))) OR (((Data[40] OR Data[1]) AND Data[32]) OR ((Data[37] OR Data[35]) AND (Data[1] AND Data[45]))))))) OR ((((Data[25] OR Data[42]) AND ((((((Data[35] XOR (NOT Data[28])) XOR (Data[12] OR Data[17])) OR Data[25]) XOR ((((Data[3] XOR Data[2]) XOR Data[25]) AND (Data[32] OR Data[9])) AND (((Data[33] AND Data[43]) XOR (NOT Data[37])) XOR (Data[28] AND Data[2])))) XOR FALSE) AND Data[30])) XOR Data[36]) XOR Data[6]))) AND (NOT (NOT Data[43])));
    OutReady := 1;
    CollectInput(RESET:=TRUE);
  END_IF;
END_PROGRAM

CONFIGURATION Config0
  RESOURCE Res0 ON PLC
    TASK task0(INTERVAL := T#20ms,PRIORITY := 0);
    PROGRAM instance0 WITH task0 : Boiler;
  END_RESOURCE
END_CONFIGURATION

(* ---- RND-EXPR_stool-idiom-aspic.st ---- *)
(*
This code implements a randomly grown symbolic expression:

!((xor(xor(IN23, !((xor(xor((xor(xor(!(!(IN13)), IN37), (xor(xor(IN23, false), false)) & IN16)) & (xor(xor(!(!(IN44)), IN15 | (IN17 & IN42)), (!(IN26)) & (IN50 & IN10))), (((!(IN24)) & (!(IN13))) | (xor(xor(!(IN18), IN17 | IN37), IN31 & IN47))) | (xor(xor(!(IN27 | IN25), IN1), (!(IN38)) | (!(IN14))))), (IN24 & ((!(IN35)) & (!(IN27)))) | IN1)) & ((xor(xor((xor(xor(IN15 & IN2, IN21 & IN50), IN40 & IN35)) | IN25, IN41 & ((IN22 & IN2) & (xor(xor(IN49, IN50), IN6)))), !((IN19 | IN19) | (xor(xor(IN43, IN43), IN10))))) | ((!(IN21)) | IN43)))), !(xor(xor(xor(xor((!(IN39)) & ((xor(xor(IN14 | IN10, IN44 | IN12), IN25 | IN15)) | ((xor(xor(IN10, IN42), IN34)) & (IN17 & IN27))), xor(xor((xor(xor(xor(xor(IN23, IN14), IN25), IN47), xor(xor(IN17, true), IN20))) | ((IN7 | IN19) & IN17), IN49), (!(IN40 | IN19)) | (xor(xor(IN5, IN6 | IN37), IN14)))), !(((xor(xor(IN35, IN39), IN4)) | IN22) & (IN23 & (IN29 | IN25)))), xor(xor(IN41 | (((xor(xor(IN14, IN35), IN3)) & (IN45 & IN20)) & ((IN5 | IN1) & (!(IN43)))), ((!(!(IN25))) | IN36) & IN21), !(xor(xor(IN50, xor(xor(IN27 | IN31, IN29), IN1 | IN47)), (xor(xor(IN48, true), IN36)) | IN38)))), xor(xor(xor(xor(IN3, (IN6 | (IN20 | IN17)) | (xor(xor(xor(xor(IN21, IN25), IN9), IN41 & IN17), IN11 | IN34))), !((xor(xor(IN26, IN39), IN3)) & true)), (!((IN13 & IN41) & (!(IN30)))) & ((!(xor(xor(IN4, IN33), IN49))) & ((!(IN34)) & (xor(xor(IN3, IN9), IN27))))), xor(xor(((!(IN5)) & (IN10 & IN48)) & (!(IN44 & IN41)), IN9), xor(xor(!(xor(xor(IN20, IN29), true)), IN17 & (!(IN29))), (!(IN37)) & (IN30 & IN43)))))))) | IN39)

*)

FUNCTION_BLOCK F_CollectInput
  VAR_IN_OUT
      Data : ARRAY[1..50] OF BOOL;
  END_VAR
  VAR_INPUT
      TICK  : BOOL := 0;
      IN1   : BOOL := 0;
      IN2   : BOOL := 0;
      IN3   : BOOL := 0;
      IN4   : BOOL := 0;
      IN5   : BOOL := 0;
      RESET : BOOL := FALSE;
  END_VAR
  VAR_OUTPUT
      Finished : BOOL;
  END_VAR
  VAR
      j    : USINT := 1;
      tock : BOOL  := 0;
  END_VAR
  IF NOT RESET AND tock = NOT TICK THEN
      Data[j]   := IN1;
      Data[j+1] := IN2;
      Data[j+2] := IN3;
      Data[j+3] := IN4;
      Data[j+4] := IN5;
      j := j + 5;
      tock := TICK;
  ELSE
      j := 1;
      tock := 0;
  END_IF;
  Finished := (j > 50);
END_FUNCTION_BLOCK

PROGRAM Boiler
  VAR
    Data  : ARRAY[1..50] OF BOOL;
    Ready : BOOL;
    CollectInput : F_CollectInput;
  END_VAR
  VAR
    TICK     AT %IX1.0 : BOOL;
    IN1      AT %IX0.3 : BOOL;
    IN2      AT %IX0.4 : BOOL;
    IN3      AT %IX0.5 : BOOL;
    IN4      AT %IX0.6 : BOOL;
    IN5      AT %IX0.7 : BOOL;
    OutReady AT %QX0.0 : BOOL := FALSE;
    FeedNext AT %QX0.1 : BOOL := FALSE;
    Out      AT %QX0.2 : BOOL;
  END_VAR
  CollectInput(TICK:=TICK, IN1:=IN1, IN2:=IN2, IN3:=IN3, IN4:=IN4, IN5:=IN5);
  Ready := CollectInput.Finished;
  FeedNext := 1;
  IF Ready THEN
    Out := (NOT (((Data[23] XOR (NOT (((((((NOT (NOT Data[13])) XOR Data[37]) XOR (((Data[23] XOR FALSE) XOR FALSE) AND Data[16])) AND (((NOT (NOT Data[44])) XOR (Data[15] OR (Data[17] AND Data[42]))) XOR ((NOT Data[26]) AND (Data[50] AND Data[10])))) XOR ((((NOT Data[24]) AND (NOT Data[13])) OR (((NOT Data[18]) XOR (Data[17] OR Data[37])) XOR (Data[31] AND Data[47]))) OR (((NOT (Data[27] OR Data[25])) XOR Data[1]) XOR ((NOT Data[38]) OR (NOT Data[14]))))) XOR ((Data[24] AND ((NOT Data[35]) AND (NOT Data[27]))) OR Data[1])) AND (((((((Data[15] AND Data[2]) XOR (Data[21] AND Data[50])) XOR (Data[40] AND Data[35])) OR Data[25]) XOR (Data[41] AND ((Data[22] AND Data[2]) AND ((Data[49] XOR Data[50]) XOR Data[6])))) XOR (NOT ((Data[19] OR Data[19]) OR ((Data[43] XOR Data[43]) XOR Data[10])))) OR ((NOT Data[21]) OR Data[43]))))) XOR (NOT ((((((NOT Data[39]) AND ((((Data[14] OR Data[10]) XOR (Data[44] OR Data[12])) XOR (Data[25] OR Data[15])) OR (((Data[10] XOR Data[42]) XOR Data[34]) AND (Data[17] AND Data[27])))) XOR (((((((Data[23] XOR Data[14]) XOR Data[25]) XOR Data[47]) XOR ((Data[17] XOR TRUE) XOR Data[20])) OR ((Data[7] OR Data[19]) AND Data[17])) XOR Data[49]) XOR ((NOT (Data[40] OR Data[19])) OR ((Data[5] XOR (Data[6] OR Data[37])) XOR Data[14])))) XOR (NOT ((((Data[35] XOR Data[39]) XOR Data[4]) OR Data[22]) AND (Data[23] AND (Data[29] OR Data[25]))))) XOR (((Data[41] OR ((((Data[14] XOR Data[35]) XOR Data[3]) AND (Data[45] AND Data[20])) AND ((Data[5] OR Data[1]) AND (NOT Data[43])))) XOR (((NOT (NOT Data[25])) OR Data[36]) AND Data[21])) XOR (NOT ((Data[50] XOR (((Data[27] OR Data[31]) XOR Data[29]) XOR (Data[1] OR Data[47]))) XOR (((Data[48] XOR TRUE) XOR Data[36]) OR Data[38]))))) XOR ((((Data[3] XOR ((Data[6] OR (Data[20] OR Data[17])) OR ((((Data[21] XOR Data[25]) XOR Data[9]) XOR (Data[41] AND Data[17])) XOR (Data[11] OR Data[34])))) XOR (NOT (((Data[26] XOR Data[39]) XOR Data[3]) AND TRUE))) XOR ((NOT ((Data[13] AND Data[41]) AND (NOT Data[30]))) AND ((NOT ((Data[4] XOR Data[33]) XOR Data[49])) AND ((NOT Data[34]) AND ((Data[3] XOR Data[9]) XOR Data[27]))))) XOR (((((NOT Data[5]) AND (Data[10] AND Data[48])) AND (NOT (Data[44] AND Data[41]))) XOR Data[9]) XOR (((NOT ((Data[20] XOR Data[29]) XOR TRUE)) XOR (Data[17] AND (NOT Data[29]))) XOR ((NOT Data[37]) AND (Data[30] AND Data[43])))))))) OR Data[39]));
    OutReady := 1;
    CollectInput(RESET:=TRUE);
  END_IF;
END_PROGRAM

CONFIGURATION Config0
  RESOURCE Res0 ON PLC
    TASK task0(INTERVAL := T#20ms,PRIORITY := 0);
    PROGRAM instance0 WITH task0 : Boiler;
  END_RESOURCE
END_CONFIGURATION

(* ---- RND-EXPR_sweat-dovey-chows.st ---- *)
(*
This code implements a randomly grown symbolic expression:

((((xor(xor(xor(xor(IN9, (IN28 | ((IN18 & IN41) & (!(IN11)))) & (!(!(IN14)))), !(IN42)), !((((!(IN37)) & (IN26 | IN33)) & (xor(xor(IN4, IN35 & IN47), IN26 | IN39))) | ((IN25 | (IN13 | IN10)) & (xor(xor(IN17 | IN24, !(IN3)), xor(xor(IN34, IN24), IN19)))))), IN14 & ((xor(xor(!(IN18 | IN24), !(!(IN12))), xor(xor(IN7 & IN41, IN16 & IN28), IN5))) & IN6))) | ((IN28 & ((xor(xor(!(!(IN13)), (IN47 | IN47) & (!(IN5))), IN48)) | (xor(xor(IN36 | (IN14 & IN16), IN29), IN5)))) & (((xor(xor(!(xor(xor(IN29, IN44), IN41)), (xor(xor(IN30, IN31), IN19)) | (!(IN1))), xor(xor(IN16 | IN45, xor(xor(IN46, IN31), IN41)), IN28 & IN20))) & (xor(xor(IN48, (!(IN28)) | (IN35 | IN45)), (!(IN16)) | (IN9 | IN38)))) | IN35))) & (!(!(IN31)))) & IN7) & (((IN11 & ((xor(xor(((xor(xor(xor(xor(IN46, IN2), IN34), xor(xor(IN1, IN46), IN5)), !(IN30))) & ((IN17 & IN13) & IN29)) | (xor(xor(IN22, IN14), (!(IN41)) & (IN33 & IN43))), !(!(xor(xor(!(IN29), !(IN14)), !(IN31))))), IN28)) & (xor(xor(IN11, (xor(xor(IN14, IN24), IN25 & (IN39 | true))) | (!(xor(xor(xor(xor(IN29, IN10), IN23), IN22 | IN34), xor(xor(IN48, IN33), IN32))))), (!(!(IN1 | IN36))) & (IN20 | IN14))))) & ((xor(xor((xor(xor(xor(xor(xor(xor(IN11, !(IN21)), xor(xor(IN38, true), true)), IN28 | (IN3 | IN25)), xor(xor(IN21 & IN47, IN6 & IN6), IN30 & IN17)), IN27), (xor(xor(!(IN15), xor(xor(IN3, IN36), IN50)), xor(xor(IN19, IN43), IN5))) & IN5)) | IN37, (IN8 | (xor(xor(!(IN50 & IN50), IN13 | (IN19 & IN12)), (IN30 | IN41) | IN46))) & (!(xor(xor((!(IN27)) & (IN11 & IN13), IN20), (IN48 | IN22) | IN6)))), (IN13 | (!(xor(xor(!(IN22), xor(xor(IN33, IN14), IN48)), IN5 | IN41)))) & (xor(xor(!(!(IN3)), (xor(xor(xor(xor(IN31, IN46), IN41), IN49 & IN30), true)) & (xor(xor(true, IN20 & IN41), !(IN13)))), xor(xor((!(IN5)) | (IN14 & IN28), xor(xor(xor(xor(IN6, IN45), IN46), xor(xor(IN30, IN20), IN4)), xor(xor(IN49, IN9), IN19))), (IN19 | IN2) | IN43))))) & (!(IN38)))) | IN48)

*)

FUNCTION_BLOCK F_CollectInput
  VAR_IN_OUT
      Data : ARRAY[1..50] OF BOOL;
  END_VAR
  VAR_INPUT
      TICK  : BOOL := 0;
      IN1   : BOOL := 0;
      IN2   : BOOL := 0;
      IN3   : BOOL := 0;
      IN4   : BOOL := 0;
      IN5   : BOOL := 0;
      RESET : BOOL := FALSE;
  END_VAR
  VAR_OUTPUT
      Finished : BOOL;
  END_VAR
  VAR
      j    : USINT := 1;
      tock : BOOL  := 0;
  END_VAR
  IF NOT RESET AND tock = NOT TICK THEN
      Data[j]   := IN1;
      Data[j+1] := IN2;
      Data[j+2] := IN3;
      Data[j+3] := IN4;
      Data[j+4] := IN5;
      j := j + 5;
      tock := TICK;
  ELSE
      j := 1;
      tock := 0;
  END_IF;
  Finished := (j > 50);
END_FUNCTION_BLOCK

PROGRAM Boiler
  VAR
    Data  : ARRAY[1..50] OF BOOL;
    Ready : BOOL;
    CollectInput : F_CollectInput;
  END_VAR
  VAR
    TICK     AT %IX1.0 : BOOL;
    IN1      AT %IX0.3 : BOOL;
    IN2      AT %IX0.4 : BOOL;
    IN3      AT %IX0.5 : BOOL;
    IN4      AT %IX0.6 : BOOL;
    IN5      AT %IX0.7 : BOOL;
    OutReady AT %QX0.0 : BOOL := FALSE;
    FeedNext AT %QX0.1 : BOOL := FALSE;
    Out      AT %QX0.2 : BOOL;
  END_VAR
  CollectInput(TICK:=TICK, IN1:=IN1, IN2:=IN2, IN3:=IN3, IN4:=IN4, IN5:=IN5);
  Ready := CollectInput.Finished;
  FeedNext := 1;
  IF Ready THEN
    Out := ((((((((Data[9] XOR ((Data[28] OR ((Data[18] AND Data[41]) AND (NOT Data[11]))) AND (NOT (NOT Data[14])))) XOR (NOT Data[42])) XOR (NOT ((((NOT Data[37]) AND (Data[26] OR Data[33])) AND ((Data[4] XOR (Data[35] AND Data[47])) XOR (Data[26] OR Data[39]))) OR ((Data[25] OR (Data[13] OR Data[10])) AND (((Data[17] OR Data[24]) XOR (NOT Data[3])) XOR ((Data[34] XOR Data[24]) XOR Data[19])))))) XOR (Data[14] AND ((((NOT (Data[18] OR Data[24])) XOR (NOT (NOT Data[12]))) XOR (((Data[7] AND Data[41]) XOR (Data[16] AND Data[28])) XOR Data[5])) AND Data[6]))) OR ((Data[28] AND ((((NOT (NOT Data[13])) XOR ((Data[47] OR Data[47]) AND (NOT Data[5]))) XOR Data[48]) OR (((Data[36] OR (Data[14] AND Data[16])) XOR Data[29]) XOR Data[5]))) AND (((((NOT ((Data[29] XOR Data[44]) XOR Data[41])) XOR (((Data[30] XOR Data[31]) XOR Data[19]) OR (NOT Data[1]))) XOR (((Data[16] OR Data[45]) XOR ((Data[46] XOR Data[31]) XOR Data[41])) XOR (Data[28] AND Data[20]))) AND ((Data[48] XOR ((NOT Data[28]) OR (Data[35] OR Data[45]))) XOR ((NOT Data[16]) OR (Data[9] OR Data[38])))) OR Data[35]))) AND (NOT (NOT Data[31]))) AND Data[7]) AND (((Data[11] AND (((((((((Data[46] XOR Data[2]) XOR Data[34]) XOR ((Data[1] XOR Data[46]) XOR Data[5])) XOR (NOT Data[30])) AND ((Data[17] AND Data[13]) AND Data[29])) OR ((Data[22] XOR Data[14]) XOR ((NOT Data[41]) AND (Data[33] AND Data[43])))) XOR (NOT (NOT (((NOT Data[29]) XOR (NOT Data[14])) XOR (NOT Data[31]))))) XOR Data[28]) AND ((Data[11] XOR (((Data[14] XOR Data[24]) XOR (Data[25] AND (Data[39] OR TRUE))) OR (NOT ((((Data[29] XOR Data[10]) XOR Data[23]) XOR (Data[22] OR Data[34])) XOR ((Data[48] XOR Data[33]) XOR Data[32]))))) XOR ((NOT (NOT (Data[1] OR Data[36]))) AND (Data[20] OR Data[14]))))) AND ((((((((((Data[11] XOR (NOT Data[21])) XOR ((Data[38] XOR TRUE) XOR TRUE)) XOR (Data[28] OR (Data[3] OR Data[25]))) XOR (((Data[21] AND Data[47]) XOR (Data[6] AND Data[6])) XOR (Data[30] AND Data[17]))) XOR Data[27]) XOR ((((NOT Data[15]) XOR ((Data[3] XOR Data[36]) XOR Data[50])) XOR ((Data[19] XOR Data[43]) XOR Data[5])) AND Data[5])) OR Data[37]) XOR ((Data[8] OR (((NOT (Data[50] AND Data[50])) XOR (Data[13] OR (Data[19] AND Data[12]))) XOR ((Data[30] OR Data[41]) OR Data[46]))) AND (NOT ((((NOT Data[27]) AND (Data[11] AND Data[13])) XOR Data[20]) XOR ((Data[48] OR Data[22]) OR Data[6]))))) XOR ((Data[13] OR (NOT (((NOT Data[22]) XOR ((Data[33] XOR Data[14]) XOR Data[48])) XOR (Data[5] OR Data[41])))) AND (((NOT (NOT Data[3])) XOR (((((Data[31] XOR Data[46]) XOR Data[41]) XOR (Data[49] AND Data[30])) XOR TRUE) AND ((TRUE XOR (Data[20] AND Data[41])) XOR (NOT Data[13])))) XOR ((((NOT Data[5]) OR (Data[14] AND Data[28])) XOR ((((Data[6] XOR Data[45]) XOR Data[46]) XOR ((Data[30] XOR Data[20]) XOR Data[4])) XOR ((Data[49] XOR Data[9]) XOR Data[19]))) XOR ((Data[19] OR Data[2]) OR Data[43]))))) AND (NOT Data[38]))) OR Data[48]));
    OutReady := 1;
    CollectInput(RESET:=TRUE);
  END_IF;
END_PROGRAM

CONFIGURATION Config0
  RESOURCE Res0 ON PLC
    TASK task0(INTERVAL := T#20ms,PRIORITY := 0);
    PROGRAM instance0 WITH task0 : Boiler;
  END_RESOURCE
END_CONFIGURATION

(* ---- RND-EXPR_swift-casus-newer.st ---- *)
(*
This code implements a randomly grown symbolic expression:

IN41 & (((!(xor(xor(true | (IN11 & (xor(xor(xor(xor(!(IN18), IN9 | IN2), IN35 | IN48), IN33), !(IN37 & IN42)))), IN23), (!(xor(xor(IN46, xor(xor(xor(xor(IN24, IN10), IN35), IN18 & IN26), IN24)), IN6))) | (!(IN40))))) | (xor(xor((!(IN24)) & (!(IN30)), !(IN4)), !(((!((IN48 & IN1) & IN29)) | (IN43 | ((IN3 | IN24) & IN26))) | (xor(xor(IN11, ((false | IN12) & (IN18 | IN46)) | (IN29 & (!(IN39)))), IN11)))))) | (!(xor(xor(IN36, IN25 | (xor(xor(false | ((xor(xor(xor(xor(IN34, IN44), IN45), IN23), IN13)) | (xor(xor(!(IN4), false | IN22), IN35 | IN35))), IN41 | (xor(xor(IN23, !(!(IN30))), IN40))), xor(xor(((IN7 | IN13) & (IN16 | IN46)) & IN24, ((IN45 | IN32) | (IN5 & IN30)) | (xor(xor(IN5, IN28), IN29 & IN13))), ((!(IN17)) | IN50) & IN28)))), !(IN45)))))

*)

FUNCTION_BLOCK F_CollectInput
  VAR_IN_OUT
      Data : ARRAY[1..50] OF BOOL;
  END_VAR
  VAR_INPUT
      TICK  : BOOL := 0;
      IN1   : BOOL := 0;
      IN2   : BOOL := 0;
      IN3   : BOOL := 0;
      IN4   : BOOL := 0;
      IN5   : BOOL := 0;
      RESET : BOOL := FALSE;
  END_VAR
  VAR_OUTPUT
      Finished : BOOL;
  END_VAR
  VAR
      j    : USINT := 1;
      tock : BOOL  := 0;
  END_VAR
  IF NOT RESET AND tock = NOT TICK THEN
      Data[j]   := IN1;
      Data[j+1] := IN2;
      Data[j+2] := IN3;
      Data[j+3] := IN4;
      Data[j+4] := IN5;
      j := j + 5;
      tock := TICK;
  ELSE
      j := 1;
      tock := 0;
  END_IF;
  Finished := (j > 50);
END_FUNCTION_BLOCK

PROGRAM Boiler
  VAR
    Data  : ARRAY[1..50] OF BOOL;
    Ready : BOOL;
    CollectInput : F_CollectInput;
  END_VAR
  VAR
    TICK     AT %IX1.0 : BOOL;
    IN1      AT %IX0.3 : BOOL;
    IN2      AT %IX0.4 : BOOL;
    IN3      AT %IX0.5 : BOOL;
    IN4      AT %IX0.6 : BOOL;
    IN5      AT %IX0.7 : BOOL;
    OutReady AT %QX0.0 : BOOL := FALSE;
    FeedNext AT %QX0.1 : BOOL := FALSE;
    Out      AT %QX0.2 : BOOL;
  END_VAR
  CollectInput(TICK:=TICK, IN1:=IN1, IN2:=IN2, IN3:=IN3, IN4:=IN4, IN5:=IN5);
  Ready := CollectInput.Finished;
  FeedNext := 1;
  IF Ready THEN
    Out := (Data[41] AND (((NOT (((TRUE OR (Data[11] AND (((((NOT Data[18]) XOR (Data[9] OR Data[2])) XOR (Data[35] OR Data[48])) XOR Data[33]) XOR (NOT (Data[37] AND Data[42]))))) XOR Data[23]) XOR ((NOT ((Data[46] XOR ((((Data[24] XOR Data[10]) XOR Data[35]) XOR (Data[18] AND Data[26])) XOR Data[24])) XOR Data[6])) OR (NOT Data[40])))) OR ((((NOT Data[24]) AND (NOT Data[30])) XOR (NOT Data[4])) XOR (NOT (((NOT ((Data[48] AND Data[1]) AND Data[29])) OR (Data[43] OR ((Data[3] OR Data[24]) AND Data[26]))) OR ((Data[11] XOR (((FALSE OR Data[12]) AND (Data[18] OR Data[46])) OR (Data[29] AND (NOT Data[39])))) XOR Data[11]))))) OR (NOT ((Data[36] XOR (Data[25] OR (((FALSE OR (((((Data[34] XOR Data[44]) XOR Data[45]) XOR Data[23]) XOR Data[13]) OR (((NOT Data[4]) XOR (FALSE OR Data[22])) XOR (Data[35] OR Data[35])))) XOR (Data[41] OR ((Data[23] XOR (NOT (NOT Data[30]))) XOR Data[40]))) XOR (((((Data[7] OR Data[13]) AND (Data[16] OR Data[46])) AND Data[24]) XOR (((Data[45] OR Data[32]) OR (Data[5] AND Data[30])) OR ((Data[5] XOR Data[28]) XOR (Data[29] AND Data[13])))) XOR (((NOT Data[17]) OR Data[50]) AND Data[28]))))) XOR (NOT Data[45])))));
    OutReady := 1;
    CollectInput(RESET:=TRUE);
  END_IF;
END_PROGRAM

CONFIGURATION Config0
  RESOURCE Res0 ON PLC
    TASK task0(INTERVAL := T#20ms,PRIORITY := 0);
    PROGRAM instance0 WITH task0 : Boiler;
  END_RESOURCE
END_CONFIGURATION

(* ---- RND-EXPR_taffy-boned-moped.st ---- *)
(*
This code implements a randomly grown symbolic expression:

xor(xor(((!(xor(xor(xor(xor(IN26 | IN7, (!(!(IN29 | IN2))) | (!(!(xor(xor(IN18, IN45), IN3))))), IN24 & IN5), xor(xor(xor(xor(!(!(IN25 | IN32)), xor(xor(xor(xor(IN6 & IN50, IN30 & IN7), IN6), (xor(xor(IN5, IN21), IN37)) & (xor(xor(IN39, IN13), IN11))), (IN34 | IN37) | (IN45 & IN2))), (IN38 | (IN23 | IN8)) | (xor(xor(true, IN31), IN12))), (xor(xor((xor(xor(IN16, IN6), IN12)) & IN14, IN41), xor(xor(!(IN27), false | IN20), IN3 & IN37))) & (!(IN36))), !(!(IN12)))), ((xor(xor(!(IN44 & IN4), (xor(xor(IN13, IN29), IN19)) & (IN27 & IN50)), IN43 | (IN27 & IN8))) | (IN6 & ((IN16 | IN42) & (IN36 & IN3)))) | (xor(xor(!(xor(xor(xor(xor(IN36, IN40), IN47), xor(xor(IN45, true), IN10)), IN46 & IN11)), !(xor(xor(xor(xor(IN2, IN40), IN47), false), IN37))), IN27 | (xor(xor(IN38 | IN39, false & IN13), IN46))))))) | ((xor(xor(IN36, (xor(xor(xor(xor((xor(xor(IN20, IN32), IN47)) | (IN47 & IN25), IN30), (xor(xor(IN43, IN32), IN26)) & (!(IN35))), !(IN45)), !(!(IN8 & IN11)))) & (IN3 & (!((!(IN48)) | (IN20 | IN48))))), IN4)) | IN37)) | (xor(xor(xor(xor(IN23, true), (((((xor(xor(IN15, IN44), IN34)) & (!(IN23))) | IN47) & (xor(xor((IN2 | IN13) & (IN12 | IN7), xor(xor(IN31 | IN21, !(IN37)), !(IN15))), (IN36 | IN17) | (!(IN23))))) & (!((xor(xor(IN46 | IN33, IN42 & IN36), IN36)) | (IN9 & (IN18 & IN29))))) & (!((xor(xor(IN38, xor(xor(IN29 | IN39, xor(xor(IN4, IN45), IN24)), !(IN20))), xor(xor(IN35, xor(xor(IN10, IN48), IN26)), !(IN32)))) | IN42))), (!(IN20)) | (((IN21 | (((xor(xor(IN49, IN5), IN1)) | (IN18 | IN10)) | (xor(xor(xor(xor(IN45, IN29), IN5), xor(xor(IN44, IN49), IN43)), IN29 | IN10)))) | (IN33 & (!(IN46)))) & (xor(xor(!(xor(xor(IN5 & (IN27 & IN27), IN46), IN47 & (xor(xor(IN32, IN23), IN49)))), IN34), !((!(IN35 & IN46)) & IN41))))), IN20)), IN42), (((IN27 | (!(!((IN21 & (IN33 | IN46)) & IN10)))) & IN17) | ((!(IN14 & IN33)) & IN23)) & (!(IN11)))

*)

FUNCTION_BLOCK F_CollectInput
  VAR_IN_OUT
      Data : ARRAY[1..50] OF BOOL;
  END_VAR
  VAR_INPUT
      TICK  : BOOL := 0;
      IN1   : BOOL := 0;
      IN2   : BOOL := 0;
      IN3   : BOOL := 0;
      IN4   : BOOL := 0;
      IN5   : BOOL := 0;
      RESET : BOOL := FALSE;
  END_VAR
  VAR_OUTPUT
      Finished : BOOL;
  END_VAR
  VAR
      j    : USINT := 1;
      tock : BOOL  := 0;
  END_VAR
  IF NOT RESET AND tock = NOT TICK THEN
      Data[j]   := IN1;
      Data[j+1] := IN2;
      Data[j+2] := IN3;
      Data[j+3] := IN4;
      Data[j+4] := IN5;
      j := j + 5;
      tock := TICK;
  ELSE
      j := 1;
      tock := 0;
  END_IF;
  Finished := (j > 50);
END_FUNCTION_BLOCK

PROGRAM Boiler
  VAR
    Data  : ARRAY[1..50] OF BOOL;
    Ready : BOOL;
    CollectInput : F_CollectInput;
  END_VAR
  VAR
    TICK     AT %IX1.0 : BOOL;
    IN1      AT %IX0.3 : BOOL;
    IN2      AT %IX0.4 : BOOL;
    IN3      AT %IX0.5 : BOOL;
    IN4      AT %IX0.6 : BOOL;
    IN5      AT %IX0.7 : BOOL;
    OutReady AT %QX0.0 : BOOL := FALSE;
    FeedNext AT %QX0.1 : BOOL := FALSE;
    Out      AT %QX0.2 : BOOL;
  END_VAR
  CollectInput(TICK:=TICK, IN1:=IN1, IN2:=IN2, IN3:=IN3, IN4:=IN4, IN5:=IN5);
  Ready := CollectInput.Finished;
  FeedNext := 1;
  IF Ready THEN
    Out := (((((NOT (((((Data[26] OR Data[7]) XOR ((NOT (NOT (Data[29] OR Data[2]))) OR (NOT (NOT ((Data[18] XOR Data[45]) XOR Data[3]))))) XOR (Data[24] AND Data[5])) XOR (((((NOT (NOT (Data[25] OR Data[32]))) XOR (((((Data[6] AND Data[50]) XOR (Data[30] AND Data[7])) XOR Data[6]) XOR (((Data[5] XOR Data[21]) XOR Data[37]) AND ((Data[39] XOR Data[13]) XOR Data[11]))) XOR ((Data[34] OR Data[37]) OR (Data[45] AND Data[2])))) XOR ((Data[38] OR (Data[23] OR Data[8])) OR ((TRUE XOR Data[31]) XOR Data[12]))) XOR ((((((Data[16] XOR Data[6]) XOR Data[12]) AND Data[14]) XOR Data[41]) XOR (((NOT Data[27]) XOR (FALSE OR Data[20])) XOR (Data[3] AND Data[37]))) AND (NOT Data[36]))) XOR (NOT (NOT Data[12])))) XOR (((((NOT (Data[44] AND Data[4])) XOR (((Data[13] XOR Data[29]) XOR Data[19]) AND (Data[27] AND Data[50]))) XOR (Data[43] OR (Data[27] AND Data[8]))) OR (Data[6] AND ((Data[16] OR Data[42]) AND (Data[36] AND Data[3])))) OR (((NOT ((((Data[36] XOR Data[40]) XOR Data[47]) XOR ((Data[45] XOR TRUE) XOR Data[10])) XOR (Data[46] AND Data[11]))) XOR (NOT ((((Data[2] XOR Data[40]) XOR Data[47]) XOR FALSE) XOR Data[37]))) XOR (Data[27] OR (((Data[38] OR Data[39]) XOR (FALSE AND Data[13])) XOR Data[46])))))) OR (((Data[36] XOR ((((((((Data[20] XOR Data[32]) XOR Data[47]) OR (Data[47] AND Data[25])) XOR Data[30]) XOR (((Data[43] XOR Data[32]) XOR Data[26]) AND (NOT Data[35]))) XOR (NOT Data[45])) XOR (NOT (NOT (Data[8] AND Data[11])))) AND (Data[3] AND (NOT ((NOT Data[48]) OR (Data[20] OR Data[48])))))) XOR Data[4]) OR Data[37])) OR ((((Data[23] XOR TRUE) XOR (((((((Data[15] XOR Data[44]) XOR Data[34]) AND (NOT Data[23])) OR Data[47]) AND ((((Data[2] OR Data[13]) AND (Data[12] OR Data[7])) XOR (((Data[31] OR Data[21]) XOR (NOT Data[37])) XOR (NOT Data[15]))) XOR ((Data[36] OR Data[17]) OR (NOT Data[23])))) AND (NOT ((((Data[46] OR Data[33]) XOR (Data[42] AND Data[36])) XOR Data[36]) OR (Data[9] AND (Data[18] AND Data[29]))))) AND (NOT (((Data[38] XOR (((Data[29] OR Data[39]) XOR ((Data[4] XOR Data[45]) XOR Data[24])) XOR (NOT Data[20]))) XOR ((Data[35] XOR ((Data[10] XOR Data[48]) XOR Data[26])) XOR (NOT Data[32]))) OR Data[42])))) XOR ((NOT Data[20]) OR (((Data[21] OR ((((Data[49] XOR Data[5]) XOR Data[1]) OR (Data[18] OR Data[10])) OR ((((Data[45] XOR Data[29]) XOR Data[5]) XOR ((Data[44] XOR Data[49]) XOR Data[43])) XOR (Data[29] OR Data[10])))) OR (Data[33] AND (NOT Data[46]))) AND (((NOT (((Data[5] AND (Data[27] AND Data[27])) XOR Data[46]) XOR (Data[47] AND ((Data[32] XOR Data[23]) XOR Data[49])))) XOR Data[34]) XOR (NOT ((NOT (Data[35] AND Data[46])) AND Data[41])))))) XOR Data[20])) XOR Data[42]) XOR ((((Data[27] OR (NOT (NOT ((Data[21] AND (Data[33] OR Data[46])) AND Data[10])))) AND Data[17]) OR ((NOT (Data[14] AND Data[33])) AND Data[23])) AND (NOT Data[11])));
    OutReady := 1;
    CollectInput(RESET:=TRUE);
  END_IF;
END_PROGRAM

CONFIGURATION Config0
  RESOURCE Res0 ON PLC
    TASK task0(INTERVAL := T#20ms,PRIORITY := 0);
    PROGRAM instance0 WITH task0 : Boiler;
  END_RESOURCE
END_CONFIGURATION

(* ---- RND-EXPR_tower-mucho-giant.st ---- *)
(*
This code implements a randomly grown symbolic expression:

(!(!(IN30))) & IN39

*)

FUNCTION_BLOCK F_CollectInput
  VAR_IN_OUT
      Data : ARRAY[1..50] OF BOOL;
  END_VAR
  VAR_INPUT
      TICK  : BOOL := 0;
      IN1   : BOOL := 0;
      IN2   : BOOL := 0;
      IN3   : BOOL := 0;
      IN4   : BOOL := 0;
      IN5   : BOOL := 0;
      RESET : BOOL := FALSE;
  END_VAR
  VAR_OUTPUT
      Finished : BOOL;
  END_VAR
  VAR
      j    : USINT := 1;
      tock : BOOL  := 0;
  END_VAR
  IF NOT RESET AND tock = NOT TICK THEN
      Data[j]   := IN1;
      Data[j+1] := IN2;
      Data[j+2] := IN3;
      Data[j+3] := IN4;
      Data[j+4] := IN5;
      j := j + 5;
      tock := TICK;
  ELSE
      j := 1;
      tock := 0;
  END_IF;
  Finished := (j > 50);
END_FUNCTION_BLOCK

PROGRAM Boiler
  VAR
    Data  : ARRAY[1..50] OF BOOL;
    Ready : BOOL;
    CollectInput : F_CollectInput;
  END_VAR
  VAR
    TICK     AT %IX1.0 : BOOL;
    IN1      AT %IX0.3 : BOOL;
    IN2      AT %IX0.4 : BOOL;
    IN3      AT %IX0.5 : BOOL;
    IN4      AT %IX0.6 : BOOL;
    IN5      AT %IX0.7 : BOOL;
    OutReady AT %QX0.0 : BOOL := FALSE;
    FeedNext AT %QX0.1 : BOOL := FALSE;
    Out      AT %QX0.2 : BOOL;
  END_VAR
  CollectInput(TICK:=TICK, IN1:=IN1, IN2:=IN2, IN3:=IN3, IN4:=IN4, IN5:=IN5);
  Ready := CollectInput.Finished;
  FeedNext := 1;
  IF Ready THEN
    Out := ((NOT (NOT Data[30])) AND Data[39]);
    OutReady := 1;
    CollectInput(RESET:=TRUE);
  END_IF;
END_PROGRAM

CONFIGURATION Config0
  RESOURCE Res0 ON PLC
    TASK task0(INTERVAL := T#20ms,PRIORITY := 0);
    PROGRAM instance0 WITH task0 : Boiler;
  END_RESOURCE
END_CONFIGURATION
